// 랙·모듈은 새 표본이 왔을 때만 다시 계산 (PLC 주기마다 300개를 계산하지 않음)
IF NOT _bCalculated OR i_stState.nSampleSeq <> _nLastSeq OR q_bValid <> _bLastValid THEN
	_bCalculated := TRUE;
	_nLastSeq := i_stState.nSampleSeq;
	_bLastValid := q_bValid;
	_nOnlineRacks := 0;
	_bInitializing := FALSE;
	_bCharging := FALSE;
	_bDischarging := FALSE;
	_nBatWarn1 := 0;
	_nBatWarn2 := 0;
	FOR _nIndex := 1 TO 5 DO _anBatFault[_nIndex] := 0; END_FOR
	FOR _nRack := 1 TO GVL_PARAM.RACKS_PER_BMS DO
		q_astRack[_nRack] := _stRackEmpty;
		q_astRack[_nRack].DeviceIndex := (i_nDeviceIndex - 1) * UINT_TO_UDINT(GVL_PARAM.RACKS_PER_BMS) + UINT_TO_UDINT(_nRack);	// 전체 랙 순번 1부터
		q_astRack[_nRack].BatIndex := i_nDeviceIndex;
		q_astRack[_nRack].ModuleCount := UINT_TO_UDINT(i_stState.nModuleCount);
		q_astRack[_nRack].Status := 1; // b0 통신에러
		FOR _nModule := 1 TO GVL_PARAM.MODULES_PER_RACK DO
			_nIndex := (_nRack - 1) * GVL_PARAM.MODULES_PER_RACK + _nModule;
			q_astModule[_nIndex] := _stModuleEmpty;
			q_astModule[_nIndex].BatIndex := i_nDeviceIndex;
			q_astModule[_nIndex].RackIndex := UINT_TO_UDINT(_nRack);
			q_astModule[_nIndex].DeviceIndex := UINT_TO_UDINT(_nModule);
		END_FOR
		IF q_bValid AND _nRack <= i_stState.nRackCount THEN
			_nAnalog := (_nRack - 1) * 4;
			_nStatus := (_nRack - 1) * 9;
			_wOperation := i_stRaw.awRackStatus[_nStatus + 1];
			// 명세 RD-BAT-01 (v2.37): 배터리 eventMap v2. 칸 하나에 BMS 워드 2개 (첫 워드 b0~, 둘째 워드 b16~), 워드 안에서는 정의된 비트만 이어 붙임
			_wSysAlarm := i_stRaw.awRackStatus[_nStatus] AND SYS_ALARM_MASK;
			_wSysWarn := i_stRaw.awRackStatus[_nStatus + 2] AND SYS_WARN_MASK;
			_wSysError := i_stRaw.awRackStatus[_nStatus + 3] AND SYS_ERROR_MASK;
			_wModError := i_stRaw.awRackStatus[_nStatus + 4] AND MODULE_ERROR_MASK;
			_wErr1 := i_stRaw.awRackStatus[_nStatus + 5];
			_wErr2 := i_stRaw.awRackStatus[_nStatus + 6] AND ERROR_CODE2_MASK;
			_wFire := i_stRaw.awRackStatus[_nStatus + 7] AND FIRE_MASK;
			_wModule := i_stRaw.awRackStatus[_nStatus + 8] AND MODULE_STATUS_MASK;
			_wLock1 := 0;
			_wLock2 := 0;
			_wSelf1 := 0;
			_wSelf2 := 0;
			IF i_stState.abDetailValid[_nRack] THEN // 랙 상세는 순서대로 나눠 읽으므로 받은 랙만
				_wLock1 := i_stRaw.aawDetail[_nRack, 11] AND LOCK1_MASK;
				_wLock2 := i_stRaw.aawDetail[_nRack, 12] AND LOCK2_MASK;
				_wSelf1 := i_stRaw.aawDetail[_nRack, 13] AND SELF1_MASK;
				_wSelf2 := i_stRaw.aawDetail[_nRack, 14] AND SELF2_MASK;
			END_IF
			q_astRack[_nRack].Warning1 := WORD_TO_UDINT(_wSysWarn) OR SHL(WORD_TO_UDINT(_wSysAlarm), 16);	// S+2 | S+0
			// 명세 RD-BAT-01 (v2.48): 경고 비트 5개는 Warning2 b0~4 (S+4 b9 → b0, S+8 b0·2·4·6 → b1~4). '워드 2개' 규칙의 예외
			q_astRack[_nRack].Warning2 := WORD_TO_UDINT(SHR(_wModError, 9) AND 16#0001)
				OR SHL(WORD_TO_UDINT(_wModule AND 16#0001), 1)
				OR SHL(WORD_TO_UDINT(SHR(_wModule, 2) AND 16#0001), 2)
				OR SHL(WORD_TO_UDINT(SHR(_wModule, 4) AND 16#0001), 3)
				OR SHL(WORD_TO_UDINT(SHR(_wModule, 6) AND 16#0001), 4);
			// S+3 | S+4 (v2.48: b0~8 → b16~24, b10 → b25. b9는 Warning2)
			q_astRack[_nRack].Fault1 := WORD_TO_UDINT(_wSysError)
				OR SHL(WORD_TO_UDINT(_wModError AND 16#01FF), 16)
				OR SHL(WORD_TO_UDINT(SHR(_wModError, 10) AND 16#0001), 25);
			// S+7 (b0 → b0, b15 → b1) | S+8 (v2.48: b1·3·5·7·8 → b16~20. 경고 b0·2·4·6은 Warning2)
			q_astRack[_nRack].Fault2 := WORD_TO_UDINT(_wFire AND 16#0001) OR SHL(WORD_TO_UDINT(SHR(_wFire, 15)), 1)
				OR SHL(WORD_TO_UDINT(SHR(_wModule, 1) AND 16#0001), 16)
				OR SHL(WORD_TO_UDINT(SHR(_wModule, 3) AND 16#0001), 17)
				OR SHL(WORD_TO_UDINT(SHR(_wModule, 5) AND 16#0001), 18)
				OR SHL(WORD_TO_UDINT(SHR(_wModule, 7) AND 16#0001), 19)
				OR SHL(WORD_TO_UDINT(SHR(_wModule, 8) AND 16#0001), 20);
			// D+11 (b0·1 → b0·1, b3 → b2, b6~11 → b3~8) | D+12 (b0·1 → b16·17, b4~15 → b18~29)
			q_astRack[_nRack].Fault3 := WORD_TO_UDINT(_wLock1 AND 16#0003)
				OR SHL(WORD_TO_UDINT(SHR(_wLock1, 3) AND 16#0001), 2)
				OR SHL(WORD_TO_UDINT(SHR(_wLock1, 6) AND 16#003F), 3)
				OR SHL(WORD_TO_UDINT(_wLock2 AND 16#0003), 16)
				OR SHL(WORD_TO_UDINT(SHR(_wLock2, 4) AND 16#0FFF), 18);
			q_astRack[_nRack].Fault4 := WORD_TO_UDINT(_wErr1) OR SHL(WORD_TO_UDINT(_wErr2), 16);			// S+5 | S+6
			// D+13 | D+14 (b0~10 → b16~26, b12~15 → b27~30)
			q_astRack[_nRack].Fault5 := WORD_TO_UDINT(_wSelf1)
				OR SHL(WORD_TO_UDINT(_wSelf2 AND 16#07FF), 16)
				OR SHL(WORD_TO_UDINT(SHR(_wSelf2, 12) AND 16#000F), 27);
			_bRackWarn := (q_astRack[_nRack].Warning1 OR q_astRack[_nRack].Warning2) <> 0;	// v2.48: Warning2 포함
			_bRackFault := (q_astRack[_nRack].Fault1 OR q_astRack[_nRack].Fault2 OR q_astRack[_nRack].Fault3
				OR q_astRack[_nRack].Fault4 OR q_astRack[_nRack].Fault5) <> 0;
			_nBatWarn1 := _nBatWarn1 OR q_astRack[_nRack].Warning1;
			_nBatWarn2 := _nBatWarn2 OR q_astRack[_nRack].Warning2;
			_anBatFault[1] := _anBatFault[1] OR q_astRack[_nRack].Fault1;
			_anBatFault[2] := _anBatFault[2] OR q_astRack[_nRack].Fault2;
			_anBatFault[3] := _anBatFault[3] OR q_astRack[_nRack].Fault3;
			_anBatFault[4] := _anBatFault[4] OR q_astRack[_nRack].Fault4;
			_anBatFault[5] := _anBatFault[5] OR q_astRack[_nRack].Fault5;
			q_astRack[_nRack].Status := 0;
			q_astRack[_nRack].Status.1 := NOT _wOperation.0; // Initializing
			q_astRack[_nRack].Status.2 := _wOperation.3; // Ready = Idle RELAY ON
			q_astRack[_nRack].Status.3 := _wOperation.1; // Charge
			q_astRack[_nRack].Status.4 := _wOperation.2; // Discharge
			q_astRack[_nRack].Status.5 := _bRackWarn; // Warning 칸 중 하나라도 0이 아님
			q_astRack[_nRack].Status.6 := _bRackFault; // Fault 칸 중 하나라도 0이 아님
			q_astRack[_nRack].Status.7 := _wOperation.1 OR _wOperation.2 OR _wOperation.3; // Online
			q_astRack[_nRack].Status.10 := (SHR(i_stState.wRackContactor, _nRack - 1) AND 1) <> 0; // 랙 컨택터 붙음 (맵 v1.4 Input 27) [2026-11-13]
			q_astRack[_nRack].DcVoltage := WORD_TO_REAL(i_stRaw.awRackAnalog[_nAnalog]) * 0.1;
			q_astRack[_nRack].DcCurrent := F_UpsSignedWord(i_stRaw.awRackAnalog[_nAnalog + 1]) * 0.1;
			q_astRack[_nRack].Soc := WORD_TO_REAL(i_stRaw.awRackAnalog[_nAnalog + 2]) * 0.1;
			q_astRack[_nRack].Soh := WORD_TO_REAL(i_stRaw.awRackAnalog[_nAnalog + 3]);
			IF q_astRack[_nRack].Status.7 THEN _nOnlineRacks := _nOnlineRacks + 1; END_IF
			_bInitializing := _bInitializing OR NOT _wOperation.0;
			_bCharging := _bCharging OR _wOperation.1;
			_bDischarging := _bDischarging OR _wOperation.2;

			// 상세 데이터: 406칸. 모듈 슬롯 0부터 설치 수만큼 사용
			IF i_stState.abDetailValid[_nRack] THEN
				q_astRack[_nRack].MaxModuleTemp := F_UpsSignedWord(i_stRaw.aawDetail[_nRack, 0]) * 0.1;
				q_astRack[_nRack].MinModuleTemp := F_UpsSignedWord(i_stRaw.aawDetail[_nRack, 1]) * 0.1;
				q_astRack[_nRack].AvgModuleTemp := F_UpsSignedWord(i_stRaw.aawDetail[_nRack, 2]) * 0.1;
				q_astRack[_nRack].MaxCellVoltage := WORD_TO_REAL(i_stRaw.aawDetail[_nRack, 3]) * 0.001;
				q_astRack[_nRack].MinCellVoltage := WORD_TO_REAL(i_stRaw.aawDetail[_nRack, 4]) * 0.001;
				q_astRack[_nRack].AvgCellVoltage := WORD_TO_REAL(i_stRaw.aawDetail[_nRack, 5]) * 0.001;
				_wCellMax := 0;
				_wCellMin := 16#FFFF;
				_fTempMax := -1.0E6;
				_fTempMin := 1.0E6;
				FOR _nModule := 1 TO MIN(i_stState.nModuleCount, GVL_PARAM.MODULES_PER_RACK) DO
					_nIndex := (_nRack - 1) * GVL_PARAM.MODULES_PER_RACK + _nModule;
					// @MAP 랙 상세 D+15+m (첫 랙 30516부터), uint16 x0.01 V. m = 모듈 번호 - 1
					q_astModule[_nIndex].ModuleVolatge1 := WORD_TO_REAL(i_stRaw.aawDetail[_nRack, 14 + _nModule]) * 0.01;
					// ModuleVolatge2/3은 BMS 맵에 없어 _stModuleEmpty의 0 유지
					_fTemp := F_UpsSignedWord(i_stRaw.aawDetail[_nRack, 31 + _nModule]) * 0.1; // 맵은 모듈당 최고 온도 1개
					q_astModule[_nIndex].ModuleTemp1 := _fTemp;
					IF _fTemp > _fTempMax THEN
						_fTempMax := _fTemp;
						q_astRack[_nRack].MaxModuleTempLocationFromModule := UINT_TO_UDINT(_nModule);
					END_IF
					IF _fTemp < _fTempMin THEN
						_fTempMin := _fTemp;
						q_astRack[_nRack].MinModuleTempLocationFromModule := UINT_TO_UDINT(_nModule);
					END_IF
					_pCell := ADR(q_astModule[_nIndex].CellVoltage1);
					FOR _nCell := 1 TO MIN(GVL_PARAM.CELLS_PER_MODULE, 20) DO	// 설치 셀 수만 (맵은 모듈당 20칸, 레코드 CellVoltage15~20은 0으로 남음)
						_wCell := i_stRaw.aawDetail[_nRack, 66 + 20 * (_nModule - 1) + _nCell - 1];
						_pCell[_nCell - 1] := WORD_TO_REAL(_wCell) * 0.001;
						IF _wCell > _wCellMax THEN
							_wCellMax := _wCell;
							q_astRack[_nRack].MaxCellVoltageLocationFromModule := UINT_TO_UDINT(_nModule);
							q_astRack[_nRack].MaxCellVoltageLocationFromCell := UINT_TO_UDINT(_nCell);
						END_IF
						IF _wCell < _wCellMin THEN
							_wCellMin := _wCell;
							q_astRack[_nRack].MinCellVoltageLocationFromModule := UINT_TO_UDINT(_nModule);
							q_astRack[_nRack].MinCellVoltageLocationFromCell := UINT_TO_UDINT(_nCell);
						END_IF
					END_FOR
				END_FOR
			END_IF
		END_IF
	END_FOR
END_IF

IF q_bValid THEN
	q_stBat.OnlineRackCount := _nOnlineRacks;
	q_stBat.Status := 0;
	q_stBat.Status.1 := _bInitializing;
	q_stBat.Status.2 := NOT _bInitializing AND _nOnlineRacks = 0; // Standby
	q_stBat.Status.3 := _nOnlineRacks > 0 AND NOT _bCharging AND NOT _bDischarging; // Ready
	q_stBat.Status.4 := _bCharging;
	q_stBat.Status.5 := _bDischarging;
	// 명세 RD-BAT-02 (v2.48): BAT Warning1·Warning2·Fault1~5 = 랙 값 OR (칸 배치는 RACK과 같음). 나머지 칸은 0
	q_stBat.Warning1 := _nBatWarn1;
	q_stBat.Warning2 := _nBatWarn2;
	q_stBat.Fault1 := _anBatFault[1];
	q_stBat.Fault2 := _anBatFault[2];
	q_stBat.Fault3 := _anBatFault[3];
	q_stBat.Fault4 := _anBatFault[4];
	q_stBat.Fault5 := _anBatFault[5];
	q_stBat.Status.6 := (_nBatWarn1 OR _nBatWarn2) <> 0;	// v2.48: Warning2 포함
	q_stBat.Status.7 := (_anBatFault[1] OR _anBatFault[2] OR _anBatFault[3] OR _anBatFault[4] OR _anBatFault[5]) <> 0;
	q_stBat.Status.9 := i_stState.bSystemLock; // Emergency = 어느 랙이든 System Lock (Level 3, 현장 해제 필요)
	q_stBat.Status.11 := i_stState.bChargeContactorClosed; // 충전 컨택터 붙음 (맵 v1.4 Input 26 b0) [2026-11-13]
	q_stBat.Status.12 := i_stState.bDischargeContactorClosed; // 방전 컨택터 붙음 (맵 v1.4 Input 26 b1) [2026-11-13]
	q_stBat.Status.13 := i_stState.wRackContactor <> 0; // 명세 RD-BAT-02 (v2.28): 랙 컨택터 닫힘 = 랙 하나라도 닫힘 (Input 27 ≠ 0, EMS 단선도 DC 컨택터)
	// b8 Balancing, b10 E-stop은 맵에 정보가 없어 항상 0 (미지원)
END_IF
// Eol, 랙 충·방전 제한, 온도 셀 위치는 맵에 없어 0. RACK b8 Precharge·b9 Balancing은 미지원이라 0.

END_FUNCTION_BLOCK

// ---- 20_Module/Ups/F_UpsSignedWord.TcPOU
FUNCTION F_UpsSignedWord : REAL
VAR_INPUT i_wRaw : WORD; END_VAR

IF i_wRaw >= 16#8000 THEN
	F_UpsSignedWord := DINT_TO_REAL(WORD_TO_DINT(i_wRaw) - 65536);
ELSE
	F_UpsSignedWord := WORD_TO_REAL(i_wRaw);
END_IF

END_FUNCTION

// ---- 20_Module/Report/FB_RptSebangUps.TcPOU
FUNCTION_BLOCK FB_RptSebangUps // UPS 계측값 → UPS 보고값
VAR_INPUT
	i_stState : ST_UpsState; // 장비 상태
	i_nDeviceIndex : UDINT; // UPS 번호
	i_nOperationMode : UDINT := 1; // 0 수동, 1 자동 (FB_UpsCommand.q_nOperationMode)
END_VAR
VAR_OUTPUT
	q_stUps : ST_UpsPublish_V1; // UPS 보고값
	q_bValid : BOOL; // 유효한 장비 데이터
END_VAR
VAR
	_stEmpty : ST_UpsPublish_V1;
	_awWarn : ARRAY[0..7] OF WORD; // 워드별 경고장 비트 (I44~I51)
	_awFault : ARRAY[0..7] OF WORD; // 워드별 중고장 비트 (I44~I51)
	_i : INT;
	_b : INT; // 워드 안 비트 번호
	_wBit : WORD;
	_nWarnPos : INT; // 다음에 채울 Warning1 비트
	_nFault1Pos : INT; // 다음에 채울 Fault1 비트
	_nFault2Pos : INT; // 다음에 채울 Fault2 비트
END_VAR
VAR CONSTANT
	// 세방 맵 v3.2 Alarm Flag 색. 순서 = I44 입력, I45 정류부, I46 BBC, I47 출력, I48 인버터, I49 바이패스, I50 STATUS1, I51 STATUS2
	WARN_MASK : ARRAY[0..7] OF WORD := [16#0700, 16#0003, 16#0007, 16#00FF, 16#0000, 16#03FF, 16#0000, 16#0701]; // 경고장(노랑)
	FAULT_MASK : ARRAY[0..7] OF WORD := [16#F8FF, 16#667C, 16#0FB8, 16#3F00, 16#803F, 16#0000, 16#0081, 16#7800]; // 중고장(주황)
	FAULT1_LAST_WORD : INT := 2; // 중고장 I44~I46 → Fault1, I47~I51 → Fault2 (회사 eventMap)
END_VAR

q_stUps := _stEmpty;
q_stUps.DeviceIndex := i_nDeviceIndex;
q_stUps.Status := 1; // b0 통신에러
q_bValid := i_stState.bValid;
IF NOT q_bValid THEN
	RETURN;
END_IF

// 명세 RD-UPS-02 (v2.20, 회사 eventMap '001.UPS 경고장비트맵'): 마스크로 거른 경고장·중고장 비트를
// 맵 워드 순서(I44→I51), 워드 안 비트 순서로 b0부터 빈칸 없이 채운다. 마스크 밖 비트(운전 상태·예약)는 버림
//   Warning1 = 경고장 30개 (I44·I45·I46·I47·I49·I51) b0~b29, Warning2·3 = 0
//   Fault1 = I44·I45·I46 중고장 30개 b0~b29, Fault2 = I47·I48·I50·I51 중고장 19개 b0~b18, Fault3 = 0
// 마스크가 바뀌면 그 뒤 비트 자리가 모두 밀리므로 eventMap도 같이 고쳐야 함
_nWarnPos := 0;
_nFault1Pos := 0;
_nFault2Pos := 0;
FOR _i := 0 TO 7 DO
	_awWarn[_i] := i_stState.awAlarmStatus[_i] AND WARN_MASK[_i];
	_awFault[_i] := i_stState.awAlarmStatus[_i] AND FAULT_MASK[_i];
	FOR _b := 0 TO 15 DO
		_wBit := SHL(WORD#1, _b);
		IF (WARN_MASK[_i] AND _wBit) <> 0 THEN
			IF (_awWarn[_i] AND _wBit) <> 0 THEN
				q_stUps.Warning1 := q_stUps.Warning1 OR SHL(UDINT#1, _nWarnPos);
			END_IF
			_nWarnPos := _nWarnPos + 1;
		END_IF
		IF (FAULT_MASK[_i] AND _wBit) <> 0 THEN
			IF _i <= FAULT1_LAST_WORD THEN
				IF (_awFault[_i] AND _wBit) <> 0 THEN
					q_stUps.Fault1 := q_stUps.Fault1 OR SHL(UDINT#1, _nFault1Pos);
				END_IF
				_nFault1Pos := _nFault1Pos + 1;
			ELSE
				IF (_awFault[_i] AND _wBit) <> 0 THEN
					q_stUps.Fault2 := q_stUps.Fault2 OR SHL(UDINT#1, _nFault2Pos);
				END_IF
				_nFault2Pos := _nFault2Pos + 1;
			END_IF
		END_IF
	END_FOR
END_FOR

// 명세 RD-UPS-01: 상태 칸 (인터페이스 08.UPS 2026-11-12). 맵 워드: I45 정류부, I46 BBC, I48 인버터, I50 STATUS1, I51 STATUS2
// 운전 모드 (2026-11-25): EMS UPS 명령 101 수동·102 자동을 반영. SystemOperationMode는 0 유지
q_stUps.SystemOperationMode := 0;
q_stUps.OperationMode := i_nOperationMode;
q_stUps.Status := 0;
q_stUps.Status.1 := (q_stUps.Warning1 OR q_stUps.Warning2 OR q_stUps.Warning3) <> 0; // 경고 있음
q_stUps.Status.2 := (q_stUps.Fault1 OR q_stUps.Fault2 OR q_stUps.Fault3) <> 0; // 고장 있음
q_stUps.Status.3 := i_stState.bEmergencyStop; // e-stop (I50 b0)
q_stUps.Status.4 := i_stState.wStatus1.13; // 충전 중 (I50 b13 Batt charg Flag)

q_stUps.UPS_ModeStatus := 0;
q_stUps.UPS_ModeStatus.0 := i_stState.nBatMode = 0; // 부동충전 (BAT Mode 값을 비트로 나눔)
q_stUps.UPS_ModeStatus.1 := i_stState.nBatMode = 1; // 균등충전
q_stUps.UPS_ModeStatus.2 := i_stState.nBatMode = 2; // 대기
q_stUps.UPS_ModeStatus.3 := i_stState.nBatMode = 3; // 주기적 방전
q_stUps.UPS_ModeStatus.4 := i_stState.nBatMode = 4; // 펄스 방전
q_stUps.UPS_ModeStatus.5 := i_stState.nBatMode = 5; // 간헐충전
q_stUps.UPS_ModeStatus.6 := i_stState.wRectAlarm.8; // 비상 방전 (I45 b8 Regen mode)
q_stUps.UPS_ModeStatus.7 := i_stState.bTemperatureEnabled; // 온도보상충전 (I51 b2, 다른 모드와 동시 가능)
q_stUps.UPS_ModeStatus.8 := i_stState.wInverterAlarm.7; // ECO 모드 (I48 b7)
q_stUps.UPS_ModeStatus.9 := i_stState.wStatus1.12; // PRLT 모드 (I50 b12)
q_stUps.UPS_ModeStatus.10 := i_stState.wStatus1.11; // Droop 모드 (I50 b11)
q_stUps.UPS_ModeStatus.11 := i_stState.wRectAlarm.15; // VSM 모드 (I45 b15)
q_stUps.UPS_ModeStatus.12 := i_stState.wRectAlarm.8; // Regen 모드 (I45 b8, b6과 같은 비트)

q_stUps.MCCB_Status := SHR(WORD_TO_UDINT(i_stState.wStatus1), 1) AND 16#3F; // I50 b1~b6 → b0~b5 (b5 Out C/B는 1이 개방)
q_stUps.MCCB_Status.6 := i_stState.wOpCode.3; // 배터리 MCCB Trip (H11 OP-CODE b3, 1 = Trip, 세방 회신 2026-11-25, 명세 RD-UPS-01 v2.50)

q_stUps.RectStatus := 0;
q_stUps.RectStatus.0 := i_stState.bRectOn; // 정류부 기동 (I45 b11)
q_stUps.RectStatus.1 := i_stState.bRectNormal; // 정류부 정상 (I45 b12)
q_stUps.RectStatus.2 := i_stState.wRectAlarm.8; // Regen (I45 b8, 비상 방전)

q_stUps.BBCStatus := 0;
q_stUps.BBCStatus.0 := i_stState.bBbcOn; // 배터리 컨버터 기동 (I46 b12)
q_stUps.BBCStatus.1 := i_stState.bBbcNormal; // 배터리 컨버터 정상 (I46 b13)

q_stUps.InverterStatus := 0;
q_stUps.InverterStatus.0 := i_stState.bInverterOn; // 인버터 기동 (I48 b6)
q_stUps.InverterStatus.1 := i_stState.bInverterNormal; // 인버터 정상 (I48 b14)
q_stUps.InverterStatus.2 := i_stState.bOnInverter; // 인버터 출력 (I48 b13)

q_stUps.BypassStatus := 0;
q_stUps.BypassStatus.0 := i_stState.bOnBypass; // 바이패스 출력 (I48 b12)

q_stUps.LineInputVoltage_R := i_stState.fInputVoltageRV;
q_stUps.LineInputVoltage_S := i_stState.fInputVoltageSV;
q_stUps.LineInputVoltage_T := i_stState.fInputVoltageTV;
q_stUps.InputFrequency := i_stState.fInputFrequencyHz;
q_stUps.InputCurrent_R := i_stState.fInputCurrentRA;
q_stUps.InputCurrent_S := i_stState.fInputCurrentSA;
q_stUps.InputCurrent_T := i_stState.fInputCurrentTA;
q_stUps.InverterVoltage_R := i_stState.fInverterVoltageRV;
q_stUps.InverterVoltage_S := i_stState.fInverterVoltageSV;
q_stUps.InverterVoltage_T := i_stState.fInverterVoltageTV;
q_stUps.InverterCurrent_R := i_stState.fInverterCurrentRA;
q_stUps.InverterCurrent_S := i_stState.fInverterCurrentSA;
q_stUps.InverterCurrent_T := i_stState.fInverterCurrentTA;
q_stUps.BypassLineVoltage_R := i_stState.fBypassVoltageRV;
q_stUps.BypassLineVoltage_S := i_stState.fBypassVoltageSV;
q_stUps.BypassLineVoltage_T := i_stState.fBypassVoltageTV;
q_stUps.BypassFrequency := i_stState.fBypassFrequencyHz;
q_stUps.LineOutputVoltage_R := i_stState.fOutputVoltageRV;
q_stUps.LineOutputVoltage_S := i_stState.fOutputVoltageSV;
q_stUps.LineOutputVoltage_T := i_stState.fOutputVoltageTV;
q_stUps.FrequencyOutput := i_stState.fOutputFrequencyHz;
q_stUps.OutputCurrent_R := i_stState.fOutputCurrentRA;
q_stUps.OutputCurrent_S := i_stState.fOutputCurrentSA;
q_stUps.OutputCurrent_T := i_stState.fOutputCurrentTA;
q_stUps.DcLinkVoltage := i_stState.fDcLinkVoltageV;
q_stUps.DcLinkVoltage_High := i_stState.fDcLinkHighVoltageV;
q_stUps.DcLinkVoltage_Low := i_stState.fDcLinkLowVoltageV;
q_stUps.BatteryVoltage := i_stState.fBatteryVoltageV;
q_stUps.BatteryCurrent := i_stState.fBatteryCurrentA;
q_stUps.MPI_A_Current := i_stState.fMpiCurrentAA;
q_stUps.MPI_B_Current := i_stState.fMpiCurrentBA;
q_stUps.MPI_C_Current := i_stState.fMpiCurrentCA;
q_stUps.InputApparentPower := i_stState.fInputApparentPowerKva;
q_stUps.OutputApparentPower := i_stState.fOutputApparentPowerKva;
q_stUps.OutputActivePower := i_stState.fOutputActivePowerKw;
q_stUps.Temp1 := i_stState.fTemperature1C;
q_stUps.Temp2 := i_stState.fTemperature2C;
q_stUps.Temp3 := i_stState.fTemperature3C;
q_stUps.Temp4 := i_stState.fTemperature4C;
q_stUps.Temp5 := i_stState.fTemperature5C;
q_stUps.Temp6 := i_stState.fBatteryRoomTemperatureC;

END_FUNCTION_BLOCK

// ---- 20_Module/Report/FB_RptLsImd1000.TcPOU
FUNCTION_BLOCK FB_RptLsImd1000		// LS IMD1000 읽은 값 → IMD 보고값 (인터페이스\22. IMD.xlsx)
(* 2026-11-09. 명세 DV-11·RD-IMD-01 (v1.8)
   Status (사용자 결정 2026-11-09, 저항이 높은 경보부터)
     b0 통신에러 = 통신 이상 또는 아직 못 읽음 (나머지 칸 0)
     b1 Pre-Warning = Pre Alarm#3 동작 (IR 210 b3, 초기값 100 kΩ)
     b2 Warning = Pre Alarm#1 OR #2 동작 (IR 210 b1·b2, 초기값 40·70 kΩ)
     b3 Fault = 자가진단 오류 (IR 209 b0~2 메모리·RTC·교정) OR Device 이상 (IR 211 b1)
     b4 Alarm = Ins. Alarm 동작 (IR 210 b0, 초기값 10 kΩ)
     b5 Internal test = Self Test 진행 중 (IR 215 = 1)
     b6 External test = 버튼·DI Self Test 입력 (IR 206 b0·b1)
   Fault1 b0 = System 연결 이상 (IR 211 b2), b1 = PE 연결 이상 (IR 211 b0)
   PreAlarmSettingValue = Pre Alarm#1 Pick-up, MainAlarmSettingValue = Ins. Alarm Pick-up (설정 영역을 못 읽었으면 0)
   DeviceErrorLocation·InsulationResistanceFaultLocation은 Bender 항목이라 0 *)
VAR_INPUT
	i_stState		: ST_LsImd1000State;	// 장비 상태 (FB_LsImd1000.q_stState)
	i_nDeviceIndex	: UDINT;				// IMD 번호 (1부터)
END_VAR
VAR_OUTPUT
	q_stImd			: ST_ImdPublish_V1;		// IMD 보고값
	q_bValid		: BOOL;					// 유효한 장비 데이터
END_VAR
VAR
	_stEmpty		: ST_ImdPublish_V1;
END_VAR

q_stImd := _stEmpty;
q_stImd.DeviceIndex := i_nDeviceIndex;
q_stImd.Status := 1;	// b0 통신에러
q_bValid := i_stState.bValid;
IF NOT q_bValid THEN
	RETURN;
END_IF

q_stImd.Status := 0;
q_stImd.Status.1 := i_stState.wAlarm.3;
q_stImd.Status.2 := i_stState.wAlarm.1 OR i_stState.wAlarm.2;
q_stImd.Status.3 := (i_stState.wSelfDiag AND 16#0007) <> 0 OR i_stState.wConnect.1;
q_stImd.Status.4 := i_stState.wAlarm.0;
q_stImd.Status.5 := i_stState.wSelfTest = 1;
q_stImd.Status.6 := i_stState.wDiState.0 OR i_stState.wDiState.1;

q_stImd.InsulationResistance := i_stState.fInsulation;
IF i_stState.bSetValid THEN
	q_stImd.PreAlarmSettingValue := i_stState.nPre1Pickup;
	q_stImd.MainAlarmSettingValue := i_stState.nInsPickup;
END_IF
q_stImd.Fault1.0 := i_stState.wConnect.2;
q_stImd.Fault1.1 := i_stState.wConnect.0;

END_FUNCTION_BLOCK

// ---- 20_Module/Report/FB_RptTempHum.TcPOU
FUNCTION_BLOCK FB_RptTempHum		// 온습도계 읽은 값 → 온도 보고값 (인터페이스\07.Temperature Sensor.xlsx, 토픽 temperature_sensor)
(* 2026-11-09. status b0 통신에러(통신 이상·값 무효면 1, 온도·습도 0). location은 설치 위치 번호
   (1 PCS실, 2 BAT실, 3 UPS실, 4 FC 컨테이너실, 5 외부) *)
VAR_INPUT
	i_stState		: ST_TempHumState;		// 장비 상태 (드라이버 q_stState)
	i_nDeviceIndex	: UDINT;				// 장치 번호 (0부터, 기존 temperature_sensor 시험 데이터와 같음)
	i_nLocation		: UDINT;				// 설치 위치
END_VAR
VAR_OUTPUT
	q_stTemp		: ST_TempPublish_V1;	// 보고값
	q_bValid		: BOOL;					// 유효한 장비 데이터
END_VAR
VAR
	_stEmpty		: ST_TempPublish_V1;
END_VAR

q_stTemp := _stEmpty;
q_stTemp.DeviceIndex := i_nDeviceIndex;
q_stTemp.location := i_nLocation;
q_stTemp.status := 1;	// b0 통신에러
q_bValid := i_stState.bValid;
IF NOT q_bValid THEN
	RETURN;
END_IF
q_stTemp.status := 0;
q_stTemp.temperature := i_stState.fTemp;
q_stTemp.humidity := i_stState.fHum;

END_FUNCTION_BLOCK

// ---- 20_Module/Driver/Esolution/FB_BmsRackCommand.TcPOU
FUNCTION_BLOCK FB_BmsRackCommand		// BMS 랙 컨택터 개별 제어: EMS 랙 명령 → 랙 선택표(BMS 40001 랙 비트) 갱신 요청
(* 2026-11-10. 명세 WR-BAT-01 (v2.5). 인터페이스 100.Command BAT CommandType 11 랙 닫기 / 12 랙 열기 (Value = 랙 번호)
   BAT 질의 Q4 답변: 랙 개별·일괄 제어 모두 지원. 일괄은 CommandType 1·2 (시스템 컨택터 40013, 기존 코어 경로)
   - 랙 선택표(비트 n-1 = 랙 n, 1 = 사용)를 기억하고, 명령마다 그 랙 비트만 바꾼 표 전체를 BMS에 쓰게 한다
   - 장비 쓰기는 하지 않는다. q_bWriteReq·q_wWriteMask를 MAIN이 보고 드라이버 M_SetRackMask를 부르고 결과를 돌려준다
   - 선택표는 PERSISTENT (i_wRestore로 시작 때 한 번 읽고, q_wMask를 MAIN이 저장). 저장값이 없으면(0) 설치된 랙 전부
   - 거절: 랙 번호 범위 밖(BadRequest), 마지막 남은 랙 열기(BadRequest: 0이면 BMS가 전 랙 사용 안 함 → 전체는 일괄 2 열기로)
   - 드라이버가 바쁘면(Busy) WRITE_TIMEOUT 동안 다시 시도. 그 밖의 거절(쓰기 막힘, 통신 불가 등)은 바로 그 결과로 끝
   - 같은 상태로 바꾸는 명령도 표 전체를 다시 씀 (BMS가 다시 켜져 표가 달라졌을 때 맞춤)
   - [2026-11-13] BMS 맵 v1.4 랙 컨택터 상태(Input 30027)를 받으면 그 실제 상태를 바탕으로 비트를 바꿈.
     40013(랙 전체 연결)으로 다 붙은 뒤 옛 선택표로 써서 다른 랙을 떼는 일을 막음. 상태가 없으면 기억한 선택표 *)
VAR_INPUT
	i_stCmd			: ST_BatRackCmd;	// EMS 랙 명령 (번호가 바뀌면 새 명령)
	i_nRackCount	: UINT;				// 설치된 랙 수 (GVL_PARAM.RACKS_PER_BMS)
	i_wRestore		: WORD;				// 처음 호출 때 한 번 읽는 저장된 선택표 (GVL_PERSIST.g_awBmsRackMask[n])
	i_bAccepted		: BOOL;				// 지난 스캔의 쓰기 요청을 드라이버가 받음 (M_SetRackMask 반환값)
	i_eDriverResult	: E_UpsResult;		// 지난 스캔 드라이버 결과 (q_eRequestResult). 요청하지 않은 스캔은 None
	i_wActual		: WORD;				// BMS 랙 컨택터 실제 상태 (q_stState.wRackContactor, 30027) [2026-11-13]
	i_bActualValid	: BOOL;				// i_wActual을 믿을 수 있음 (q_stState.bContactorFeedbackKnown)
END_VAR
VAR_OUTPUT
	q_wMask			: WORD;				// 지금 선택표 (드라이버가 받은 값). MAIN이 GVL_PERSIST에 씀
	q_bMaskChanged	: BOOL;				// 이 스캔에 q_wMask가 바뀜 (PERSISTENT 바로 저장 요청)
	q_bWriteReq		: BOOL;				// 드라이버에 쓰기 요청 중
	q_wWriteMask	: WORD;				// 쓸 선택표
	q_eResult		: E_UpsResult;		// 마지막 명령 결과
	q_nLastSeq		: UDINT;			// 마지막으로 처리한 명령 번호
END_VAR
VAR
	_bInit			: BOOL;
	_wInstalled		: WORD;
	_wNew			: WORD;
	_wOld			: WORD;
	_wBase			: WORD;				// 바꿀 바탕 (실제 상태 또는 기억한 선택표)
	_tonWait		: TON;
END_VAR
VAR CONSTANT
	WRITE_TIMEOUT	: TIME := T#5S;		// 드라이버가 바쁠 때 다시 시도하는 시간
END_VAR

q_bMaskChanged := FALSE;
_wInstalled := SHL(WORD#1, MIN(i_nRackCount, 16)) - 1;
IF NOT _bInit THEN
	q_wMask := i_wRestore AND _wInstalled;
	IF q_wMask = 0 THEN
		q_wMask := _wInstalled;	// 저장값 없음 → 설치된 랙 전부
	END_IF
	_bInit := TRUE;
END_IF
_wOld := q_wMask;

// 1) 지난 스캔 쓰기 요청의 결과
IF q_bWriteReq THEN
	_tonWait(IN := TRUE, PT := WRITE_TIMEOUT);
	IF i_bAccepted THEN
		q_wMask := q_wWriteMask;
		q_eResult := E_UpsResult.Accepted;
		q_bWriteReq := FALSE;
	ELSIF i_eDriverResult <> E_UpsResult.None AND i_eDriverResult <> E_UpsResult.Busy THEN
		q_eResult := i_eDriverResult;	// 쓰기 막힘, 통신 불가, 설정 오류 등
		q_bWriteReq := FALSE;
	ELSIF _tonWait.Q THEN
		q_eResult := E_UpsResult.Busy;	// 계속 바빠서 포기
		q_bWriteReq := FALSE;
	END_IF
	IF NOT q_bWriteReq THEN
		_tonWait(IN := FALSE);
	END_IF
END_IF

// 2) 새 명령 (처리 중인 요청이 있으면 그것을 버리고 새 명령으로)
IF i_stCmd.nSeq <> q_nLastSeq AND i_stCmd.nSeq <> 0 THEN
	q_nLastSeq := i_stCmd.nSeq;
	q_bWriteReq := FALSE;
	_tonWait(IN := FALSE);
	IF i_stCmd.nRack < 1 OR i_stCmd.nRack > i_nRackCount OR i_stCmd.nRack > 16 THEN
		q_eResult := E_UpsResult.BadRequest;
	ELSE
		IF i_bActualValid THEN
			_wBase := i_wActual AND _wInstalled;	// 실제 상태 바탕
		ELSE
			_wBase := q_wMask;
		END_IF
		IF i_stCmd.bClose THEN
			_wNew := _wBase OR SHL(WORD#1, i_stCmd.nRack - 1);
		ELSE
			_wNew := _wBase AND NOT SHL(WORD#1, i_stCmd.nRack - 1);
		END_IF
		IF _wNew = 0 THEN
			q_eResult := E_UpsResult.BadRequest;	// 마지막 랙: 전체 열기는 일괄 명령(2)으로
		ELSE
			q_wWriteMask := _wNew;
			q_bWriteReq := TRUE;
			q_eResult := E_UpsResult.None;	// 처리 중
		END_IF
	END_IF
END_IF

q_bMaskChanged := q_wMask <> _wOld;

END_FUNCTION_BLOCK

// ---- 20_Module/Driver/Esolution/FB_BmsContactorCommand.TcPOU
FUNCTION_BLOCK FB_BmsContactorCommand		// BMS 컨택터 하나씩 제어: EMS 명령 번호 5~10 → 드라이버 M_SetControl 요청
(* 2026-11-13. 인터페이스 100.Command BAT CommandType 5~10, BMS 맵 v1.4 Holding 40013~40015
   5 시스템(랙 전체 40013) 연결   6 시스템 차단
   7 충전 컨택터(40014) 닫기      8 충전 컨택터 열기
   9 방전 컨택터(40015) 닫기      10 방전 컨택터 열기
   3 비상정지 (40012 Emergency Shutdown = 1). 2026-11-23 명세 v2.33: 코어(F_BatCmdAllowed)가 지령원 EStop을 거절해 이쪽으로 옮김
   4 초기화 (40031 Reset System = 1, 비상차단 해제). 2026-11-23 명세 v2.34 (O-19 A)
   - 장비 쓰기는 하지 않는다. q_bWriteReq·q_eControl·q_bOn을 MAIN이 보고 드라이버 M_SetControl을 부르고 결과를 돌려준다
   - 3~10 밖이면 BadRequest. 드라이버가 바쁘면(Busy) WRITE_TIMEOUT 동안 다시 시도. 그 밖의 거절(쓰기 막힘, 통신 불가 등)은 바로 그 결과로 끝
   - 코어 순서(유닛 정지 확인)는 거치지 않는다 (랙 개별 11·12와 같음). 일괄 투입·개방은 1·2 (코어 경로) *)
VAR_INPUT
	i_stCmd			: ST_BatCtlCmd;		// EMS 명령 (번호가 바뀌면 새 명령)
	i_bAccepted		: BOOL;				// 지난 스캔의 쓰기 요청을 드라이버가 받음 (M_SetControl 반환값)
	i_eDriverResult	: E_UpsResult;		// 지난 스캔 드라이버 결과 (q_eRequestResult). 요청하지 않은 스캔은 None
END_VAR
VAR_OUTPUT
	q_bWriteReq		: BOOL;				// 드라이버에 쓰기 요청 중
	q_eControl		: E_EsolutionControl;	// 쓸 컨택터
	q_bOn			: BOOL;				// TRUE = 닫기(붙이기), FALSE = 열기(떼기)
	q_eResult		: E_UpsResult;		// 마지막 명령 결과
	q_nLastSeq		: UDINT;			// 마지막으로 처리한 명령 번호
END_VAR
VAR
	_tonWait		: TON;
END_VAR
VAR CONSTANT
	WRITE_TIMEOUT	: TIME := T#5S;		// 드라이버가 바쁠 때 다시 시도하는 시간
END_VAR

// 1) 지난 스캔 쓰기 요청의 결과
IF q_bWriteReq THEN
	_tonWait(IN := TRUE, PT := WRITE_TIMEOUT);
	IF i_bAccepted THEN
		q_eResult := E_UpsResult.Accepted;
		q_bWriteReq := FALSE;
	ELSIF i_eDriverResult <> E_UpsResult.None AND i_eDriverResult <> E_UpsResult.Busy THEN
		q_eResult := i_eDriverResult;	// 쓰기 막힘, 통신 불가 등
		q_bWriteReq := FALSE;
	ELSIF _tonWait.Q THEN
		q_eResult := E_UpsResult.Busy;	// 계속 바빠서 포기
		q_bWriteReq := FALSE;
	END_IF
	IF NOT q_bWriteReq THEN
		_tonWait(IN := FALSE);
	END_IF
END_IF

// 2) 새 명령 (처리 중인 요청이 있으면 그것을 버리고 새 명령으로)
IF i_stCmd.nSeq <> q_nLastSeq AND i_stCmd.nSeq <> 0 THEN
	q_nLastSeq := i_stCmd.nSeq;
	q_bWriteReq := FALSE;
	_tonWait(IN := FALSE);
	q_eResult := E_UpsResult.None;	// 처리 중
	CASE i_stCmd.nType OF
		3:		q_eControl := E_EsolutionControl.EmergencyShutdown;
		4:		q_eControl := E_EsolutionControl.ResetSystem;
		5, 6:	q_eControl := E_EsolutionControl.SystemContactor;
		7, 8:	q_eControl := E_EsolutionControl.ChargeContactor;
		9, 10:	q_eControl := E_EsolutionControl.DischargeContactor;
	ELSE
		q_eResult := E_UpsResult.BadRequest;
	END_CASE
	IF q_eResult = E_UpsResult.None THEN
		q_bOn := (i_stCmd.nType MOD 2) = 1 OR i_stCmd.nType = 4;	// 3 비상정지·4 초기화 = 켜기(1), 5·7·9 = 닫기
		q_bWriteReq := TRUE;
	END_IF
END_IF

END_FUNCTION_BLOCK

// ---- 20_Module/Ups/FB_UpsSafetyResponse.TcPOU
FUNCTION_BLOCK FB_UpsSafetyResponse		// 사고·고장 대응 동작 (C안): 원인 → UPS·BMS 명령, 될 때까지 2초마다 다시 보내고 10초 넘으면 오류 표시
(* 2026-11-17. 명세 SQ-05 (v2.16), 동작시퀀스 7쪽 표. 기반 없음(신규).
   변경: 2026-11-18 ESD(b12) 대응을 나눔: 바이패스 절체 빼고 인버터 정지(H105) 추가, 순서 기다리지 않고 연달아 보냄 (명세 v2.18)
   변경: 2026-11-20 화재(b11)는 ESD처럼: 바이패스 절체 안 함, 인버터·BBC·정류부를 기다리지 않고 연달아 (명세 SQ-05 v2.31)
   변경: 2026-11-20 바이패스 이상(UPS Warning1 b16~25 = I49)이고 아직 바이패스가 아니면 바이패스 절체를 보내지 않음 → q_bBypassBlocked (v2.31, O-17)
   변경: 2026-11-20 세방 맵 '인버터정지 To Bypass': 출력·인버터 중고장, 화재, MBS C/B Fail(대응 원인 b13)은 바이패스 절체가
         확인된 뒤 인버터 정지(H105)도 보냄. 절체가 확인 안 되면 인버터를 끄지 않음(부하 유지). 원인은 q_nRespCause (명세 SQ-05 v2.30)
   변경: 2026-11-18 "3초 확인·최대 3번 → 실패로 멈춤"을 "될 때까지 2초마다 계속 보냄, 10초 넘게 안 되면 오류 표시(그 뒤에도 계속)"로 바꿈 (명세 v2.19, 데스틴 PCS 통신 방식)
   - 원인은 FB_UpsSafetyStage.q_nRespCause (지금 걸린 대응 원인, v2.30). 여러 원인이면 동작을 합친다
   - 동작 6개 (비트): 0 충전 컨택터 열기(BMS 40014=0), 1 BMS 컨택터 전부 열기(40013~15=0),
     2 바이패스 절체(UPS H109), 3 BBC 정지(H107), 4 정류부 정지(H103), 5 인버터 정지(H105, ESD 또는 절체 확인 뒤)
   - 먼저 확인해서 이미 그 상태면 명령하지 않는다. 명령 → i_tResend 기다림 → 안 됐으면 다시. 될 때까지 계속
   - i_tFail 넘게 안 되면 q_wFailed(오류)를 켠다. 오류가 켜져도 계속 보낸다. 되면 오류는 꺼진다
   - 드라이버가 못 받은 명령(바쁨·통신 끊김)은 기다리지 않고 다음 스캔에 다시 보낸다 (보낸 횟수에 넣지 않음)
   - 된 동작은 원인이 사라졌다가 다시 생길 때까지 다시 하지 않는다 (사람이 다시 켠 것을 되돌리지 않음)
   - UPS 명령은 스캔마다 하나. 순서는 바이패스 → 인버터(절체 확인 뒤) → BBC → 정류부: 앞 동작이 되거나 오류가 켜져야 다음 동작을 보낸다
     BMS는 전부 열기가 필요하면 충전만 열기는 하지 않는다
   - ESD나 화재가 걸려 있으면: 바이패스 절체는 하지 않는다(다른 원인이 요구해도). UPS 명령은 앞 동작을 기다리지 않고
     인버터 → BBC → 정류부 순으로 연달아 보낸다
   - i_bEnable(전체 스위치 AND 쓰기 관문)이 꺼지면 모두 처음 상태로
   - UPS 명령은 i_ipUps로 직접 보낸다. BMS 명령은 q_eBmsReq(그 스캔만)로 내고 MAIN이 드라이버를 부른다
   - 복귀(다시 켜기), MCCB Trip, 바이패스 포함 출력 차단, BMS E-stop은 하지 않는다
   변경: 2026-11-25 이중화 절체 때 상대의 된 동작 기억을 이어받음 (명세 RED-01·SQ-05 v2.49): i_bInheritLoad 때 i_wInheritDone을 담아 두고,
         그 동작이 필요해지면 보내지 않고 '됨'으로 둠 (사람이 다시 켠 것을 되돌리지 않음). 쓰기 허가·UPS 읽기 뒤 i_tInheritSettle 동안 안 쓰인 비트와
         i_tInheritMax가 지난 비트는 버림 *)
VAR_INPUT
	i_bEnable		: BOOL;					// GVL_PERSIST.g_bUpsSafetyRespEnable AND 장비 쓰기 관문
	i_nCause		: UDINT;				// FB_UpsSafetyStage.q_nRespCause (대응 원인, v2.30)
	i_stUps			: ST_UpsPublish_V1;		// UPS 보고값 (RectStatus b0, BBCStatus b0, InverterStatus b0, BypassStatus b0)
	i_bUpsValid		: BOOL;					// UPS 통신 정상
	i_stBms			: ST_EsolutionState;	// BMS 상태 (컨택터 30026·30027)
	i_ipUps			: I_Ups;				// UPS 명령 대상
	i_tResend		: TIME := T#2S;			// 보낸 뒤 다시 보내기까지 (응답 대기 1초 + 쉼 1초)
	i_tFail			: TIME := T#10S;		// 이 시간 넘게 안 되면 오류 표시 (보내기는 계속)
	i_bInheritLoad	: BOOL;					// 이 스캔에 이어받을 기억을 담음 (이중화: 이 PLC가 Active가 되는 순간, 명세 RED-01 v2.49)
	i_wInheritDone	: WORD;					// 이어받을 된 동작 비트 (대기 중 받은 상대의 q_wDone)
	i_tInheritSettle: TIME := T#3S;			// 쓰기 허가 + UPS 읽기 뒤 이 시간 동안 필요해지지 않은 이어받은 비트는 버림
	i_tInheritMax	: TIME := T#30S;		// 이어받은 비트는 담은 뒤 이 시간이 지나면 버림
END_VAR
VAR_OUTPUT
	q_wNeeded		: WORD;					// 지금 필요한 동작 (비트 0~5)
	q_wDone			: WORD;					// 된 동작
	q_wFailed		: WORD;					// 오류: i_tFail 넘게 안 된 동작 (계속 보내는 중. EMS 칸 없음, PLC 안에서만)
	q_eBmsReq		: UINT;					// BMS 요청: 0 없음, 1 충전 컨택터 열기, 2 전부 열기 (MAIN이 드라이버에 전달)
	q_nBmsSeq		: UDINT;				// 전부 열기 명령 번호 (M_SetStateCmd 중복 거르기용, 16#7F000000부터)
	q_anTry			: ARRAY[0..5] OF UINT;	// 동작별 보낸 횟수 (드라이버가 받은 것만, 65535에서 멈춤)
	q_bEsd			: BOOL;					// ESD·화재 대응 중 (순서 기다리지 않음, 바이패스 절체 안 함, v2.31 화재 포함)
	q_bBypassBlocked : BOOL;				// 바이패스 이상이라 바이패스 절체를 보내지 않는 중 (기록 BypassBlocked, v2.31)
	q_wInherit		: WORD;					// 아직 쓰지 않은 이어받은 된 동작 비트 (v2.49)
END_VAR
VAR
	_anState		: ARRAY[0..5] OF UINT;	// 0 보낼 차례, 1 보낸 뒤 기다림, 2 됨
	_atonResend		: ARRAY[0..5] OF TON;
	_atonFail		: ARRAY[0..5] OF TON;
	_abAchieved		: ARRAY[0..5] OF BOOL;
	_k				: INT;
	_i				: INT;
	_bNeed			: BOOL;
	_bUpsSent		: BOOL;					// 이번 스캔에 UPS 명령을 이미 시도함
	_bUpsHold		: BOOL;					// 앞 UPS 동작이 진행 중이라 뒤 동작은 기다림 (ESD가 아닐 때)
	_nBmsCount		: UDINT;
	_wBit			: WORD;
	_eCmd			: E_UpsCommand;
	_bInvStopArmed	: BOOL;					// 인버터 정지 To Bypass: 바이패스가 확인돼 인버터 정지를 시작함 (원인이 사라질 때까지 유지)
	_wInherit		: WORD;					// 이어받은 된 동작 비트 (쓰거나 버리면 지움, v2.49)
	_tonInheritSettle : TON;
	_tonInheritMax	: TON;
END_VAR
VAR CONSTANT
	ACT_CHG_OPEN	: INT := 0;
	ACT_BMS_OPEN	: INT := 1;
	ACT_BYPASS		: INT := 2;
	ACT_BBC_OFF		: INT := 3;
	ACT_RECT_OFF	: INT := 4;
	ACT_INV_OFF		: INT := 5;
	// 진행 순서 (동작 번호). UPS는 바이패스 → 인버터 → BBC → 정류부
	ORDER			: ARRAY[0..5] OF INT := [0, 1, 2, 5, 3, 4];
	// SQ-01 원인 비트
	C_BMS_MINOR		: UDINT := 16#00000004;	// b2
	C_BBC_GROUP		: UDINT := 16#00000388;	// b3 BMS Major, b7 지락(RCD)1, b8 BBC 중고장, b9 지락(RCD)2
	C_RECT			: UDINT := 16#00000010;	// b4 입력·정류부 중고장
	C_INV			: UDINT := 16#00002060;	// b5 출력, b6 인버터 중고장, b13 MBS C/B Fail → 바이패스 절체
	C_INV_STOP		: UDINT := 16#00002460;	// b5, b6, b13 MBS: 맵 '인버터정지 To Bypass', b10 BMS Level 3: 7쪽 표 5단계 '인버터 정지/바이패스 절체' (v2.54) → 절체 확인 뒤 인버터 정지 (화재는 v2.31부터 ESD처럼)
	C_FULL			: UDINT := 16#00000400;	// b10 BMS Level 3 (화재는 v2.31부터 C_ESD)
	C_ESD			: UDINT := 16#00001800;	// b11 화재, b12 ESD: 바이패스 절체 안 함, 인버터·BBC·정류부 정지 + BMS 전부 열기 (v2.31)
	W1_BYPASS		: UDINT := 16#03FF0000;	// UPS Warning1 b16~25 = I49 바이패스 이상 (맵 'To Bypass 절체 안 됨')
	BMS_SEQ_BASE	: UDINT := 16#7F000000;
END_VAR

// 이중화 이어받기 (명세 RED-01·SQ-05 v2.49): 담고, 오래되면 버림
IF i_bInheritLoad THEN
	_wInherit := i_wInheritDone AND 16#003F;
	_tonInheritSettle(IN := FALSE);
	_tonInheritMax(IN := FALSE);
END_IF
_tonInheritSettle(IN := _wInherit <> 0 AND i_bEnable AND i_bUpsValid, PT := i_tInheritSettle);
_tonInheritMax(IN := _wInherit <> 0, PT := i_tInheritMax);
IF _tonInheritSettle.Q OR _tonInheritMax.Q THEN
	_wInherit := 0;
END_IF

// 0) 됐는지 (확인 신호를 믿을 수 없으면 안 된 것으로 봄)
_abAchieved[ACT_CHG_OPEN] := i_stBms.bContactorFeedbackKnown AND NOT i_stBms.bChargeContactorClosed;
_abAchieved[ACT_BMS_OPEN] := i_stBms.bContactorFeedbackKnown AND i_stBms.wSystemContactor = 0 AND i_stBms.wRackContactor = 0;
_abAchieved[ACT_BYPASS] := i_bUpsValid AND i_stUps.BypassStatus.0;
_abAchieved[ACT_BBC_OFF] := i_bUpsValid AND NOT i_stUps.BBCStatus.0;
_abAchieved[ACT_RECT_OFF] := i_bUpsValid AND NOT i_stUps.RectStatus.0;
_abAchieved[ACT_INV_OFF] := i_bUpsValid AND NOT i_stUps.InverterStatus.0;

// 1) 원인 → 필요한 동작
q_wNeeded := 0;
q_bBypassBlocked := FALSE;
q_bEsd := i_bEnable AND (i_nCause AND C_ESD) <> 0;
IF i_bEnable THEN
	IF (i_nCause AND C_BMS_MINOR) <> 0 THEN q_wNeeded := q_wNeeded OR SHL(WORD#1, ACT_CHG_OPEN); END_IF
	IF (i_nCause AND C_BBC_GROUP) <> 0 THEN q_wNeeded := q_wNeeded OR SHL(WORD#1, ACT_BBC_OFF); END_IF
	IF (i_nCause AND C_RECT) <> 0 THEN
		q_wNeeded := q_wNeeded OR SHL(WORD#1, ACT_RECT_OFF) OR SHL(WORD#1, ACT_CHG_OPEN);
	END_IF
	IF (i_nCause AND C_INV) <> 0 THEN q_wNeeded := q_wNeeded OR SHL(WORD#1, ACT_BYPASS); END_IF
	IF (i_nCause AND C_FULL) <> 0 THEN
		q_wNeeded := q_wNeeded OR SHL(WORD#1, ACT_BYPASS) OR SHL(WORD#1, ACT_BBC_OFF) OR SHL(WORD#1, ACT_RECT_OFF) OR SHL(WORD#1, ACT_BMS_OPEN);
	END_IF
	// 인버터 정지 To Bypass (v2.30): 바이패스가 확인된 뒤에만 시작. 시작하면 원인이 사라질 때까지 유지
	IF (i_nCause AND C_INV_STOP) = 0 THEN
		_bInvStopArmed := FALSE;
	ELSIF _abAchieved[ACT_BYPASS] OR (_wInherit AND SHL(WORD#1, ACT_INV_OFF)) <> 0 THEN	// v2.49: 인버터 정지를 이어받으면 바이패스 확인을 기다리지 않음
		_bInvStopArmed := TRUE;
	END_IF
	IF _bInvStopArmed THEN q_wNeeded := q_wNeeded OR SHL(WORD#1, ACT_INV_OFF); END_IF
	// 바이패스 이상 (v2.31, O-17): 아직 바이패스가 아니면 절체를 보내지 않음 (부하는 인버터로 유지). 바이패스가 정상이 되면 다시 필요해짐
	IF NOT q_bEsd AND (q_wNeeded AND SHL(WORD#1, ACT_BYPASS)) <> 0 AND NOT _abAchieved[ACT_BYPASS]
		AND i_bUpsValid AND (i_stUps.Warning1 AND W1_BYPASS) <> 0 THEN
		q_bBypassBlocked := TRUE;
		q_wNeeded := q_wNeeded AND NOT SHL(WORD#1, ACT_BYPASS);
	END_IF
	IF q_bEsd THEN
		q_wNeeded := q_wNeeded OR SHL(WORD#1, ACT_INV_OFF) OR SHL(WORD#1, ACT_BBC_OFF) OR SHL(WORD#1, ACT_RECT_OFF) OR SHL(WORD#1, ACT_BMS_OPEN);
		q_wNeeded := q_wNeeded AND NOT SHL(WORD#1, ACT_BYPASS);	// 비상정지 중에 부하를 바이패스로 다시 살리지 않음
	END_IF
	IF (q_wNeeded AND SHL(WORD#1, ACT_BMS_OPEN)) <> 0 THEN
		q_wNeeded := q_wNeeded AND NOT SHL(WORD#1, ACT_CHG_OPEN);	// 전부 열기가 충전 열기를 포함
	END_IF
ELSE
	_bInvStopArmed := FALSE;
END_IF

// 2) 동작별 진행 (ORDER 순서)
_bUpsSent := FALSE;
_bUpsHold := FALSE;
q_eBmsReq := 0;
FOR _k := 0 TO 5 DO
	_i := ORDER[_k];
	_wBit := SHL(WORD#1, _i);
	_bNeed := (q_wNeeded AND _wBit) <> 0;
	_atonResend[_i](IN := _bNeed AND _anState[_i] = 1, PT := i_tResend);
	IF NOT _bNeed THEN
		_anState[_i] := 0;		// 원인이 사라짐 (또는 꺼짐) → 다음에 다시 생기면 처음부터
		q_anTry[_i] := 0;
	ELSE
		CASE _anState[_i] OF
			0:	// 보낼 차례
				IF (_wInherit AND _wBit) <> 0 THEN
					_anState[_i] := 2;	// 상대가 이미 한 동작 (이중화 이어받기, v2.49): 다시 보내지 않음
					_wInherit := _wInherit AND NOT _wBit;
				ELSIF _abAchieved[_i] THEN
					_anState[_i] := 2;	// 이미 그 상태
				ELSIF _i = ACT_CHG_OPEN OR _i = ACT_BMS_OPEN THEN
					IF q_eBmsReq = 0 THEN
						IF _i = ACT_BMS_OPEN THEN
							q_eBmsReq := 2;
							_nBmsCount := _nBmsCount + 1;
							q_nBmsSeq := BMS_SEQ_BASE + (_nBmsCount AND 16#00FFFFFF);
						ELSE
							q_eBmsReq := 1;
						END_IF
						IF q_anTry[_i] < 65535 THEN q_anTry[_i] := q_anTry[_i] + 1; END_IF
						_anState[_i] := 1;
					END_IF
				ELSIF NOT _bUpsSent AND NOT _bUpsHold AND i_ipUps <> 0 THEN
					CASE _i OF
						ACT_BYPASS:		_eCmd := E_UpsCommand.ToBypass;
						ACT_BBC_OFF:	_eCmd := E_UpsCommand.BbcOff;
						ACT_RECT_OFF:	_eCmd := E_UpsCommand.RectifierOff;
						ACT_INV_OFF:	_eCmd := E_UpsCommand.InverterOff;
					END_CASE
					_bUpsSent := TRUE;	// UPS는 스캔마다 하나
					IF i_ipUps.M_RequestCommand(_eCmd) THEN
						IF q_anTry[_i] < 65535 THEN q_anTry[_i] := q_anTry[_i] + 1; END_IF
						_anState[_i] := 1;
					END_IF	// 못 받았으면 0에 남아 다음 스캔에 다시
				END_IF
			1:	// 보낸 뒤 기다림
				IF _abAchieved[_i] THEN
					_anState[_i] := 2;
				ELSIF _atonResend[_i].Q THEN
					_anState[_i] := 0;	// 다시 보냄
				END_IF
		END_CASE
	END_IF
	_atonFail[_i](IN := _bNeed AND _anState[_i] <> 2, PT := i_tFail);
	// ESD가 아니면 앞 UPS 동작이 되거나 오류가 켜질 때까지 뒤 UPS 동작은 기다림
	IF _i >= ACT_BYPASS AND _bNeed AND _anState[_i] <> 2 AND NOT _atonFail[_i].Q AND NOT q_bEsd THEN
		_bUpsHold := TRUE;
	END_IF
END_FOR

q_wDone := 0;
q_wFailed := 0;
FOR _i := 0 TO 5 DO
	IF _anState[_i] = 2 THEN q_wDone := q_wDone OR SHL(WORD#1, _i); END_IF
	IF _atonFail[_i].Q THEN q_wFailed := q_wFailed OR SHL(WORD#1, _i); END_IF
END_FOR
q_wInherit := _wInherit;

END_FUNCTION_BLOCK

// ---- 20_Module/Ups/FB_UpsSafetyStage.TcPOU
(* LiB-UPS 사고·고장 단계 판정 (④보호 표시 / 장치: UPS·BAT). 2026-11-05.
   기반 없음(신규). 동작시퀀스 7쪽(이솔루션 2026-10-23) 단계표를 따른다.
   변경: 2026-11-09 UPS 경고·고장 4번 칸을 없앰. STATUS 비트를 Warning3 하위·Fault3 상위에서 읽음 (명세 RD-UPS-02 v1.6)
   변경: 2026-11-18 UPS 경고·고장 칸을 회사 eventMap 순서로 읽음 (Warning1·Fault1·Fault2, 명세 RD-UPS-02 v2.20)
   변경: 2026-11-18 기록(FB_UpsSafetyLog)용 출력 q_nLatched·q_bAckPulse·q_nAckCleared 추가 (명세 SQ-01 v2.21). 판정은 그대로
   변경: 2026-11-20 대응(SQ-05)용 원인 q_nRespCause 추가 (명세 SQ-05 v2.30, 세방 맵 Alarm Flag 비트별 동작). 단계 판정은 그대로
         - b4: '기동 안 됨' 2비트(Fault1 b7 입력 상회전, b18 Pre Magnet Fail) 뺌
         - b5: 출력 과전류 R/S/T(Fault2 b0~2)는 i_tOutOcDelay(15분) 계속될 때만, 출력 과전류 Trip(b3~5)은 바로
         - b8: 배터리 과전류(Fault1 b23)는 i_tBattOcDelay(10분) 계속될 때만, 나머지 BBC 중고장은 바로
         - b13: MBS C/B Fail(Fault2 b14, I50 b7). 단계 없음, 대응만
   변경: 2026-11-23 Fault(4~6단계)도 원인이 풀리면 바로 내림. 확인 전 유지(래치)와 i_bAck·q_bAckPending·q_nLatched·q_bAckPulse·q_nAckCleared 없앰
         (명세 SQ-01 v2.38: 확인은 EMS가 하므로 PMS에 확인 신호가 오지 않아, 붙잡은 Fault가 재시작 전까지 안 풀렸음)
   변경: 2026-11-23 i_bClear 추가: 이중화 대기 중에는 원인을 비움 (명세 RED-02 v2.45: 장비를 읽지 않으니 마지막 값이 옛 값. 넘겨받는 순간 옛 값으로 대응하지 않게)
   부호·단위: 해당 없음. 명세: C:\gil\UPS\명세작업\UPS_명세서.md SQ-01, SQ-05
   차단·정지는 UPS(UMS)와 BMS가 스스로 한다. 이 FB는 판정과 표시만 하고 장비에 아무것도 쓰지 않는다. *)
FUNCTION_BLOCK FB_UpsSafetyStage
VAR_INPUT
	i_stUps			: ST_UpsPublish_V1;	// UPS 보고값 (FB_RptSebangUps.q_stUps)
	i_bUpsValid		: BOOL;				// UPS 데이터 유효 (통신 정상)
	i_stBat			: ST_BatPublish_V1;	// 짝 BAT 보고값 (FB_RptEsolutionBat.q_stBat)
	i_bBatValid		: BOOL;				// BAT 데이터 유효 (통신 정상)
	i_tOutOcDelay	: TIME := T#15M;	// 출력 과전류 R/S/T가 이만큼 계속되면 대응 (세방 맵 '15분후 인버터정지 To Bypass', SQ-05 v2.30)
	i_bClear		: BOOL;				// 원인을 비움 (이중화 대기 중, 명세 RED-02 v2.45). 통신 끊김 때 마지막 값 유지보다 우선
	i_tBattOcDelay	: TIME := T#10M;	// 배터리 과전류가 이만큼 계속되면 대응 (세방 맵 '10분후 정지', SQ-05 v2.30)
END_VAR
VAR_OUTPUT
	q_nStage		: UINT;				// 대표 단계 0~6 (걸린 단계 중 가장 높은 것)
	q_wStageMask	: WORD;				// 걸린 단계 목록. bit n = n단계 (n = 1~6). 높은 순서로 모두 표시할 때 사용
	q_nCause		: UDINT;			// 원인 비트 (아래 CAUSE_* 표). q_nActiveCause와 같음 (v2.38: Fault도 붙잡지 않음)
	q_nActiveCause	: UDINT;			// 지금 실제로 걸린 원인만
	q_bUpsCommFault	: BOOL;				// UPS 통신장애 (단계와 별도 상태). 끊긴 동안 UPS 원인은 마지막 값을 유지
	q_bBatCommFault	: BOOL;				// BAT 통신장애 (단계와 별도 상태). 끊긴 동안 BAT 원인은 마지막 값을 유지
	q_nRespCause	: UDINT;			// 대응(FB_UpsSafetyResponse)용 원인. 비트 배치는 q_nActiveCause와 같고 b13 MBS C/B Fail 추가 (SQ-05 v2.30)
END_VAR
VAR
	_nUpsCause		: UDINT;			// UPS에서 나온 원인 (통신이 끊기면 마지막 값 유지)
	_nBatCause		: UDINT;			// BAT에서 나온 원인 (통신이 끊기면 마지막 값 유지)
	_nUpsResp		: UDINT;			// UPS에서 나온 대응 원인 (통신이 끊기면 마지막 값 유지)
	_tonOutOc		: TON;				// 출력 과전류 R/S/T 지속
	_tonBattOc		: TON;				// 배터리 과전류 지속
	_i				: INT;
END_VAR
VAR CONSTANT
	(* 원인 비트 → 단계. 순서 = 비트 번호 *)
	CAUSE_STAGE		: ARRAY[0..12] OF UINT := [
		1,	// b0  AC·DC SPD (I51 b8·b9)
		1,	// b1  UPS 경고장 (SPD·BMS Minor 제외)
		2,	// b2  BMS Minor (I51 b10)
		3,	// b3  BMS Major (I51 b11)
		3,	// b4  UPS 입력·정류부 중고장 (I44·I45)
		3,	// b5  UPS 출력 중고장 (I47)
		3,	// b6  UPS 인버터 중고장 (I48)
		3,	// b7  배터리 DC 전로 지락(RCD) 1단계 (I51 b12, 명세 v2.50 세방 회신)
		4,	// b8  배터리 컨버터(BBC) 중고장 (I46)
		4,	// b9  배터리 DC 전로 지락(RCD) 2단계 (I51 b13, 명세 v2.50 세방 회신)
		5,	// b10 BMS Level 3 (BAT Status b9 System Lock)
		5,	// b11 화재 (I51 b14)
		6];	// b12 ESD (I50 b0)
	(* UPS 보고 칸 안의 비트 (명세 RD-UPS-02 v2.20, 회사 eventMap 순서) *)
	W1_SPD			: UDINT := 16#18000000;	// Warning1 b27 AC SPD (I51 b8), b28 DC SPD (I51 b9)
	W1_BMS_MINOR	: UDINT := 16#20000000;	// Warning1 b29 BMS Minor (I51 b10)
	F1_INPUT		: UDINT := 16#003FFFFF;	// Fault1 b0~b21 입력·정류부 (I44·I45)
	F1_BBC			: UDINT := 16#3FC00000;	// Fault1 b22~b29 배터리 컨버터 (I46)
	F2_OUTPUT		: UDINT := 16#0000003F;	// Fault2 b0~b5 출력 (I47)
	F2_INVERTER		: UDINT := 16#00001FC0;	// Fault2 b6~b12 인버터 (I48)
	F2_ESD			: UDINT := 16#00002000;	// Fault2 b13 Emergency Stop (I50 b0). b14 MBS C/B Fail (I50 b7)은 단계 없음
	F2_BMS_MAJOR	: UDINT := 16#00008000;	// Fault2 b15 BMS Major (I51 b11)
	F2_RCD1			: UDINT := 16#00010000;	// Fault2 b16 지락(RCD) 1단계 (I51 b12)
	F2_RCD2			: UDINT := 16#00020000;	// Fault2 b17 지락(RCD) 2단계 (I51 b13)
	F2_FIRE			: UDINT := 16#00040000;	// Fault2 b18 화재 (I51 b14)
	(* 대응 원인 (SQ-05 v2.30, 세방 맵 Alarm Flag 정류부·배터리컨버터·인버터 칸) *)
	F1_START_BLOCK	: UDINT := 16#00040080;	// Fault1 b7 입력 상회전 (I44 b7), b18 Pre Magnet Fail (I45 b9): 맵 '기동 안 됨' → 명령 없음
	F1_BATT_OC		: UDINT := 16#00800000;	// Fault1 b23 배터리 과전류 (I46 b4): 맵 '10분후 정지'
	F2_OUT_OC		: UDINT := 16#00000007;	// Fault2 b0~2 출력 과전류 R/S/T (I47 b8~10): 맵 '15분후 인버터정지 To Bypass'
	F2_MBS			: UDINT := 16#00004000;	// Fault2 b14 MBS C/B Fail (I50 b7): 맵 '인버터정지 To Bypass', 단계 없음
	RESP_MBS		: UDINT := 16#00002000;	// 대응 원인 b13 MBS C/B Fail
END_VAR

// 1) UPS 원인. 통신이 끊기면 마지막 값을 그대로 둔다 (단계를 내리지 않음)
q_bUpsCommFault := NOT i_bUpsValid;
IF i_bUpsValid THEN
	_nUpsCause := 0;
	IF (i_stUps.Warning1 AND W1_SPD) <> 0 THEN _nUpsCause := _nUpsCause OR 16#0001; END_IF
	IF ((i_stUps.Warning1 AND NOT (W1_SPD OR W1_BMS_MINOR)) OR i_stUps.Warning2 OR i_stUps.Warning3) <> 0 THEN _nUpsCause := _nUpsCause OR 16#0002; END_IF
	IF (i_stUps.Warning1 AND W1_BMS_MINOR) <> 0 THEN _nUpsCause := _nUpsCause OR 16#0004; END_IF
	IF (i_stUps.Fault2 AND F2_BMS_MAJOR) <> 0 THEN _nUpsCause := _nUpsCause OR 16#0008; END_IF
	IF (i_stUps.Fault1 AND F1_INPUT) <> 0 THEN _nUpsCause := _nUpsCause OR 16#0010; END_IF
	IF (i_stUps.Fault2 AND F2_OUTPUT) <> 0 THEN _nUpsCause := _nUpsCause OR 16#0020; END_IF
	IF (i_stUps.Fault2 AND F2_INVERTER) <> 0 THEN _nUpsCause := _nUpsCause OR 16#0040; END_IF
	IF (i_stUps.Fault2 AND F2_RCD1) <> 0 THEN _nUpsCause := _nUpsCause OR 16#0080; END_IF
	IF (i_stUps.Fault1 AND F1_BBC) <> 0 THEN _nUpsCause := _nUpsCause OR 16#0100; END_IF
	IF (i_stUps.Fault2 AND F2_RCD2) <> 0 THEN _nUpsCause := _nUpsCause OR 16#0200; END_IF
	IF (i_stUps.Fault2 AND F2_FIRE) <> 0 THEN _nUpsCause := _nUpsCause OR 16#0800; END_IF
	IF (i_stUps.Fault2 AND F2_ESD) <> 0 THEN _nUpsCause := _nUpsCause OR 16#1000; END_IF
	// 대응 원인 (SQ-05 v2.30): 단계 원인에서 b4·b5·b8을 맵 동작 기준으로 다시 정하고 b13을 더함
	_tonOutOc(IN := (i_stUps.Fault2 AND F2_OUT_OC) <> 0, PT := i_tOutOcDelay);
	_tonBattOc(IN := (i_stUps.Fault1 AND F1_BATT_OC) <> 0, PT := i_tBattOcDelay);
	_nUpsResp := _nUpsCause AND NOT UDINT#16#00000130;
	IF (i_stUps.Fault1 AND F1_INPUT AND NOT F1_START_BLOCK) <> 0 THEN _nUpsResp := _nUpsResp OR 16#0010; END_IF
	IF (i_stUps.Fault2 AND F2_OUTPUT AND NOT F2_OUT_OC) <> 0 OR _tonOutOc.Q THEN _nUpsResp := _nUpsResp OR 16#0020; END_IF
	IF (i_stUps.Fault1 AND F1_BBC AND NOT F1_BATT_OC) <> 0 OR _tonBattOc.Q THEN _nUpsResp := _nUpsResp OR 16#0100; END_IF
	IF (i_stUps.Fault2 AND F2_MBS) <> 0 THEN _nUpsResp := _nUpsResp OR RESP_MBS; END_IF
END_IF

// 2) BAT 원인
q_bBatCommFault := NOT i_bBatValid;
IF i_bBatValid THEN
	_nBatCause := 0;
	IF i_stBat.Status.9 THEN _nBatCause := _nBatCause OR 16#0400; END_IF	// BMS Level 3 (System Lock)
END_IF

// 이중화 대기 중: 원인과 지연 타이머를 비움 (명세 RED-02 v2.45)
IF i_bClear THEN
	_nUpsCause := 0;
	_nBatCause := 0;
	_nUpsResp := 0;
	_tonOutOc(IN := FALSE, PT := i_tOutOcDelay);
	_tonBattOc(IN := FALSE, PT := i_tBattOcDelay);
END_IF
q_nActiveCause := _nUpsCause OR _nBatCause;
q_nRespCause := _nUpsResp OR _nBatCause;

// 3) Warning·Fault 모두 원인이 풀리면 바로 내림 (v2.38. 확인은 EMS가 함). 통신이 끊긴 장비 원인은 위에서 마지막 값 유지
q_nCause := q_nActiveCause;

// 4) 단계 목록과 대표 단계
q_wStageMask := 0;
q_nStage := 0;
FOR _i := 0 TO 12 DO
	IF (q_nCause AND SHL(UDINT#1, _i)) <> 0 THEN
		q_wStageMask := q_wStageMask OR SHL(WORD#1, CAUSE_STAGE[_i]);
		q_nStage := MAX(q_nStage, CAUSE_STAGE[_i]);
	END_IF
END_FOR

END_FUNCTION_BLOCK

// ---- 20_Module/Ups/FB_UpsSafetyLog.TcPOU
FUNCTION_BLOCK FB_UpsSafetyLog		// UPS 사고·고장 단계 기록: FB_UpsSafetyStage 결과를 PMS 이벤트 로그에 남김 (EMS로는 안 보냄)
(* 사고·고장 단계·원인 기록 (④보호 표시 / 장치: UPS·BAT). 2026-11-18.
   기반: 예전 작업본 pms-standard-main FB_UpsSafetyLog (2026-11-09, 명세 v2.0). 저장소 밖 C:\gil\UPS_보관\pms-standard-main
   변경: UPSstd로 옮김. 기록은 PMS 이벤트 로그(TwinCAT 이벤트 로거, XAE Error List)에만. 이벤트 클래스 PmsUps는
     로거 리스너(FB_MqttLoggerListener)가 받지 않아 EMS(pms_log)로 가지 않는다 (명세 SQ-01 v2.21).
     시험용 출력 q_bSettled 등과 안정 시간 입력 i_tSettle을 더함.
   변경: 2026-11-19 대응 동작(FB_UpsSafetyResponse) 기록 추가: 처음 보낸 명령, 완료, 10초 오류 (명세 SQ-01·SQ-05 v2.22)
   변경: 2026-11-23 확인 대기(AckPending)·Fault 확인(FaultAck) 기록 없앰. PMS 안에서 Fault를 붙잡지 않음 (명세 SQ-01 v2.38)
   부호·단위: 해당 없음. 명세: C:\gil\UPS\명세작업\UPS_명세서.md SQ-01 "기록"
   - 원인 알람(CauseActive): 원인 비트마다 발생·해소 1회 ("UPS n 사고·고장 k단계: 원인"). 심각도 1~3단계 Warning, 4~5 Error, 6 Critical
   - 단계 바뀜(StageChange): 대표 단계가 바뀔 때마다 메시지 1회
   - 통신장애(CommLost): 한 번이라도 통신이 됐던 장비가 끊겼을 때만 알람 (설치 안 된 장비는 기록 안 함)
   - 대응 명령(RespCmd): 동작을 처음 보낼 때 1번. 2초마다 다시 보내는 것은 남기지 않음 (보낸 횟수 0 → 1 이상)
   - 대응 완료(RespDone): 동작이 될 때 1번 (보낸 횟수, 보내기 전에 이미 그 상태였으면 그렇게)
   - 대응 오류(RespFail): 10초 넘게 안 된 동작마다 알람. 되거나 필요 없어지면 해소
   - 바이패스 절체 안 함(BypassBlocked): 바이패스 이상이라 절체를 보내지 않는 동안 알람 (명세 SQ-05 v2.31, 2026-11-20)
   - 켜진 뒤 i_tSettle 동안은 기록하지 않음 (부팅 직후 통신이 붙기 전 값으로 기록하지 않기 위해)
   판정은 하지 않는다. 원인 비트 순서·단계는 FB_UpsSafetyStage.CAUSE_STAGE와 같아야 한다 *)
VAR_INPUT
	i_nUps			: UINT;					// UPS 번호 (1~)
	i_nStage		: UINT;					// FB_UpsSafetyStage.q_nStage
	i_nActiveCause	: UDINT;				// FB_UpsSafetyStage.q_nActiveCause
	i_bUpsCommFault	: BOOL;					// FB_UpsSafetyStage.q_bUpsCommFault
	i_bBatCommFault	: BOOL;					// FB_UpsSafetyStage.q_bBatCommFault
	i_wRespNeeded	: WORD;					// FB_UpsSafetyResponse.q_wNeeded (지금 필요한 동작, 비트 0~5)
	i_wRespDone		: WORD;					// FB_UpsSafetyResponse.q_wDone
	i_wRespFailed	: WORD;					// FB_UpsSafetyResponse.q_wFailed (10초 넘게 안 된 동작)
	i_anRespTry		: ARRAY[0..5] OF UINT;	// FB_UpsSafetyResponse.q_anTry (동작별 보낸 횟수)
	i_bBypassBlocked : BOOL;				// FB_UpsSafetyResponse.q_bBypassBlocked (v2.31)
	i_tSettle		: TIME := T#15S;		// 켜진 뒤 기록하지 않는 시간
END_VAR
VAR_OUTPUT
	q_bSettled		: BOOL;					// 기록 시작함 (i_tSettle 지남)
	q_nRaised		: UDINT;				// 원인 알람이 발생 중인 원인 비트
	q_bUpsCommRaised : BOOL;				// UPS 통신장애 알람 발생 중
	q_bBatCommRaised : BOOL;				// BMS 통신장애 알람 발생 중
	q_nStageMsg		: UDINT;				// 단계 바뀜 메시지 보낸 수
	q_nRespCmdMsg	: UDINT;				// 대응 명령 메시지 보낸 수
	q_nRespDoneMsg	: UDINT;				// 대응 완료 메시지 보낸 수
	q_wRespFailRaised : WORD;				// 대응 오류 알람이 발생 중인 동작 비트
	q_bBypassBlockedRaised : BOOL;			// 바이패스 절체 안 함 알람 발생 중
END_VAR
VAR
	_tonSettle		: TON;
	_afbCause		: ARRAY[0..12] OF FB_LogAlarm;
	_fbUpsComm		: FB_LogAlarm;
	_fbBatComm		: FB_LogAlarm;
	_fbStage		: FB_LogMsg;
	_bUpsEverOk		: BOOL;
	_bBatEverOk		: BOOL;
	_nLastStage		: UINT;
	_asArg			: ARRAY[1..6] OF WSTRING(63);
	_stEntry		: TcEventEntry;
	_i				: INT;
	_bActive		: BOOL;
	_afbRespFail	: ARRAY[0..5] OF FB_LogAlarm;
	_fbRespCmd		: FB_LogMsg;
	_fbRespDone		: FB_LogMsg;
	_fbBypassBlocked : FB_LogAlarm;
	_wSent			: WORD;					// 한 번이라도 보낸 동작 (보낸 횟수 > 0)
	_wSentLast		: WORD;
	_wDone			: WORD;					// 필요하고 된 동작
	_wDoneLast		: WORD;
	_wBit			: WORD;
END_VAR
VAR CONSTANT
	CAUSE_STAGE		: ARRAY[0..12] OF UINT := [1, 1, 2, 3, 3, 3, 3, 3, 4, 4, 5, 5, 6];	// FB_UpsSafetyStage와 같음
	CAUSE_NAME		: ARRAY[0..12] OF WSTRING(31) := [
		"SPD", "UPS 경고장", "BMS Minor", "BMS Major", "입력·정류부 중고장", "출력 중고장", "인버터 중고장",
		"지락(RCD) 1단계", "배터리 컨버터 중고장", "지락(RCD) 2단계", "BMS Level 3", "화재", "ESD"];
	(* 대응 동작 이름 = FB_UpsSafetyResponse 동작 번호 순서 (명세 SQ-05) *)
	RESP_NAME		: ARRAY[0..5] OF WSTRING(39) := [
		"충전 컨택터 열기(BMS 40014=0)", "BMS 컨택터 전부 열기(40013~15=0)", "바이패스 절체(H109)",
		"BBC 정지(H107)", "정류부 정지(H103)", "인버터 정지(H105)"];
END_VAR

IF NOT i_bUpsCommFault THEN _bUpsEverOk := TRUE; END_IF
IF NOT i_bBatCommFault THEN _bBatEverOk := TRUE; END_IF
_tonSettle(IN := TRUE, PT := i_tSettle);
q_bSettled := _tonSettle.Q;
_wSent := 0;
FOR _i := 0 TO 5 DO
	IF i_anRespTry[_i] > 0 THEN _wSent := _wSent OR SHL(WORD#1, _i); END_IF
END_FOR
_wDone := i_wRespDone AND i_wRespNeeded;
IF NOT q_bSettled THEN
	_nLastStage := i_nStage;
	_wSentLast := _wSent;
	_wDoneLast := _wDone;
	RETURN;
END_IF

// 1) 원인 알람 (지금 실제로 걸린 원인)
q_nRaised := 0;
FOR _i := 0 TO 12 DO
	_bActive := (i_nActiveCause AND SHL(UDINT#1, _i)) <> 0;
	IF _bActive <> _afbCause[_i].q_bRaised THEN
		_asArg[1] := TO_WSTRING(i_nUps);
		_asArg[2] := TO_WSTRING(CAUSE_STAGE[_i]);
		_asArg[3] := CAUSE_NAME[_i];
	END_IF
	_stEntry := TC_EVENTS.PmsUps.CauseActive;
	IF CAUSE_STAGE[_i] >= 6 THEN
		_stEntry.eSeverity := TcEventSeverity.Critical;
	ELSIF CAUSE_STAGE[_i] >= 4 THEN
		_stEntry.eSeverity := TcEventSeverity.Error;
	ELSE
		_stEntry.eSeverity := TcEventSeverity.Warning;
	END_IF
	_afbCause[_i](i_stEntry := _stEntry, i_bActive := _bActive, i_nArgs := 3, i_asArg := _asArg);
	IF _afbCause[_i].q_bRaised THEN
		q_nRaised := q_nRaised OR SHL(UDINT#1, _i);
	END_IF
END_FOR

// 2) 대표 단계 바뀜
_fbStage(i_stEntry := TC_EVENTS.PmsUps.StageChange);
IF i_nStage <> _nLastStage THEN
	_asArg[1] := TO_WSTRING(i_nUps);
	_asArg[2] := TO_WSTRING(_nLastStage);
	_asArg[3] := TO_WSTRING(i_nStage);
	_fbStage.M_SendEvent(i_nArgs := 3, i_asArg := _asArg);
	_nLastStage := i_nStage;
	q_nStageMsg := q_nStageMsg + 1;
END_IF

// 3) 통신장애 (한 번이라도 됐던 장비만)
_bActive := i_bUpsCommFault AND _bUpsEverOk;
IF _bActive <> _fbUpsComm.q_bRaised THEN
	_asArg[1] := TO_WSTRING(i_nUps);
	_asArg[2] := "UPS";
END_IF
_fbUpsComm(i_stEntry := TC_EVENTS.PmsUps.CommLost, i_bActive := _bActive, i_nArgs := 2, i_asArg := _asArg);
q_bUpsCommRaised := _fbUpsComm.q_bRaised;
_bActive := i_bBatCommFault AND _bBatEverOk;
IF _bActive <> _fbBatComm.q_bRaised THEN
	_asArg[1] := TO_WSTRING(i_nUps);
	_asArg[2] := "BMS";
END_IF
_fbBatComm(i_stEntry := TC_EVENTS.PmsUps.CommLost, i_bActive := _bActive, i_nArgs := 2, i_asArg := _asArg);
q_bBatCommRaised := _fbBatComm.q_bRaised;

// 4) 대응 동작 (명세 SQ-05 기록, v2.22): 처음 보낸 명령, 완료, 10초 오류
_fbRespCmd(i_stEntry := TC_EVENTS.PmsUps.RespCmd);
_fbRespDone(i_stEntry := TC_EVENTS.PmsUps.RespDone);
q_wRespFailRaised := 0;
FOR _i := 0 TO 5 DO
	_wBit := SHL(WORD#1, _i);
	IF (_wSent AND _wBit) <> 0 AND (_wSentLast AND _wBit) = 0 THEN
		_asArg[1] := TO_WSTRING(i_nUps);
		_asArg[2] := RESP_NAME[_i];
		_fbRespCmd.M_SendEvent(i_nArgs := 2, i_asArg := _asArg);
		q_nRespCmdMsg := q_nRespCmdMsg + 1;
	END_IF
	IF (_wDone AND _wBit) <> 0 AND (_wDoneLast AND _wBit) = 0 THEN
		_asArg[1] := TO_WSTRING(i_nUps);
		_asArg[2] := RESP_NAME[_i];
		IF i_anRespTry[_i] = 0 THEN
			_asArg[3] := "이미 그 상태였음";
		ELSE
			_asArg[3] := WCONCAT("보낸 횟수 ", TO_WSTRING(i_anRespTry[_i]));
		END_IF
		_fbRespDone.M_SendEvent(i_nArgs := 3, i_asArg := _asArg);
		q_nRespDoneMsg := q_nRespDoneMsg + 1;
	END_IF
	_bActive := (i_wRespFailed AND _wBit) <> 0;
	IF _bActive <> _afbRespFail[_i].q_bRaised THEN
		_asArg[1] := TO_WSTRING(i_nUps);
		_asArg[2] := RESP_NAME[_i];
	END_IF
	_afbRespFail[_i](i_stEntry := TC_EVENTS.PmsUps.RespFail, i_bActive := _bActive, i_nArgs := 2, i_asArg := _asArg);
	IF _afbRespFail[_i].q_bRaised THEN
		q_wRespFailRaised := q_wRespFailRaised OR _wBit;
	END_IF
END_FOR
// 바이패스 이상이라 절체 안 함 (v2.31)
IF i_bBypassBlocked <> _fbBypassBlocked.q_bRaised THEN
	_asArg[1] := TO_WSTRING(i_nUps);
END_IF
_fbBypassBlocked(i_stEntry := TC_EVENTS.PmsUps.BypassBlocked, i_bActive := i_bBypassBlocked, i_nArgs := 1, i_asArg := _asArg);
q_bBypassBlockedRaised := _fbBypassBlocked.q_bRaised;
_wSentLast := _wSent;
_wDoneLast := _wDone;

END_FUNCTION_BLOCK

// ---- 20_Module/Mqtt/FB_EmsConfigApply.TcPOU
FUNCTION_BLOCK FB_EmsConfigApply		// EMS config(pcs·bat) → 운영 설정 (PlcTask. MAIN 액션 A_PassEmsCfg가 부름) [9-21 수정 2026-11-04: 추가]
(* - 입력 i_stCfg는 MAIN이 GVL_IF.g_stEmsCfg에서 일관되게 복사해 넘김. PCS·BMS 칸마다 번호(anPcsSeq·anBatSeq)가 바뀌면 새 레코드
   - [21번 수정 2026-11-09] is_available = 0인 값은 기본값으로 반영 (원래: 바꾸지 않고 기존 값 유지 → EMS가 한도를 풀 수 없었음)
       pcs 충전·방전 한도 0 → 그 방향 정격 (= 제한 없음). 두 방향 모두 0 → 그 PCS 유닛의 사용자 P 한도 끔 (bPEnable FALSE, 값은 ±정격)
       bat SOC 하한 0 → 0 %, 상한 0 → 100 % (감발 폭 fBand·재개 마진은 HMI 설정 그대로)
   - [UPS 2026-11-10] UPS 현장의 config/bat 레코드는 103.Config BAT UPS_V1 형식 (SocMin·SocMax = REAL, is_available 없음. UPS_MQTT_INTERFACE.md).
       그래서 bat 값은 받은 BMS(_abBatRx)만 계산에 넣고 항상 '있음'으로 봄. 아직 못 받은 BMS는 기본값(0 %·100 %)과 같아 결과에 영향 없음. pcs 쪽은 STD 그대로
   - pcs: 충전·방전 전력 한도 (kW) → 사용자 한도 stUnitLimit. 그 PCS의 유닛들에 정격 비율로 나눔, 충전은 fPMin (−). PvMarginRate는 쓰지 않음 (사양 대기)
   - bat: SOC 최소·최대 (%) → SOC 정책 stSocLimit. 배터리 그룹 전체 한 세트라 받은 BMS 값(기본값 포함) 중 가장 엄격한 값 (하한 = 가장 큰 값, 상한 = 가장 작은 값)
   - 범위 검사를 먼저 하고 통과한 값만 씀 (SOC는 FB_SocLimit.M_CheckSet과 같은 F_SocLimitSetErr). 버리면 q_bRejected (이벤트 로그 '잘못된 설정 값')
   - 쓴 값은 GVL_PERSIST라 재시작 뒤에도 남음. 설정 보호(FB_SettingGuard)가 한 번 더 지킴. 바꾸면 q_bApplied (이벤트 로그 '운영 설정 바뀜')
   - protection(배터리·배터리실 온도·습도 경고·고장)은 반영하지 않음 (값의 뜻·센서 대기. echo만)
   - M_BuildEcho: 설정 보호 뒤 실제 설정 → q_stEcho (MAIN이 GVL_IF.g_stEmsCfgEcho에 씀 → config echo) *)
VAR_INPUT
	i_bValid		: BOOL;			// 이번 스캔에 i_stCfg를 일관되게 복사함
	i_stCfg			: ST_IfEmsCfg;
	i_astUnitCfg	: ARRAY[1..GVL_PARAM.UNIT_COUNT] OF ST_UnitCfg;	// 유닛 ← PCS 번호, 정격
END_VAR
VAR_IN_OUT
	iq_stSocLimit	: ST_SocLimitSet;	// GVL_PERSIST.g_stModuleSet.stSocLimit
	iq_stUnitLimit	: ST_UnitLimitSet;	// GVL_PERSIST.g_stModuleSet.stUnitLimit
END_VAR
VAR_OUTPUT
	q_bApplied		: BOOL;			// 이번 스캔에 설정을 바꿈 (1스캔)
	q_sApplied		: WSTRING(63);
	q_bRejected		: BOOL;			// 이번 스캔에 받은 값을 버림 (1스캔)
	q_sRejected		: WSTRING(63);	// 마지막으로 버린 값과 이유
	q_nApplied		: UDINT;
	q_nRejected		: UDINT;
	q_stEcho		: ST_IfEmsCfgEcho;
END_VAR
VAR CONSTANT
	MAX_KW			: REAL := 1.0E6;	// kW. 이보다 큰 한도는 이상값
	SOC_MIN_DEFAULT	: REAL := 0.0;		// %, bat SocMin is_available 0일 때 [21번 수정 2026-11-09: 추가]
	SOC_MAX_DEFAULT	: REAL := 100.0;	// %, bat SocMax is_available 0일 때
END_VAR
VAR
	_stCfg			: ST_IfEmsCfg;		// 마지막으로 일관되게 받은 칸 (echo의 PvMarginRate)
	_anPcsSeq		: ARRAY[1..GVL_PARAM.PCS_COUNT] OF UDINT;
	_anBatSeq		: ARRAY[1..GVL_PARAM.BMS_COUNT] OF UDINT;
	_astBat			: ARRAY[1..GVL_PARAM.BMS_COUNT] OF ST_BatConfig_Rx;	// BMS마다 받아 둔 레코드 (가장 엄격한 SOC 계산)
	_astBatBefore	: ARRAY[1..GVL_PARAM.BMS_COUNT] OF ST_BatConfig_Rx;
	_abBatRx		: ARRAY[1..GVL_PARAM.BMS_COUNT] OF BOOL;	// [UPS] 그 BMS 레코드를 한 번이라도 받아 둠 (REAL 형식이라 빈 칸을 is_available로 못 가림)
	_abBatRxBefore	: ARRAY[1..GVL_PARAM.BMS_COUNT] OF BOOL;
	_stUnit			: ST_UnitLimitSet;
	_stSoc			: ST_SocLimitSet;
	_sErr			: WSTRING(63);
	p				: UINT;
	u				: UINT;
	b				: UINT;
	fSum			: REAL;
	fCh				: REAL;
	fDis			: REAL;
	fMin			: REAL;
	fMax			: REAL;
	bCh				: BOOL;
	bDis			: BOOL;
	bAny			: BOOL;
	bNewBat			: BOOL;
	bBad			: BOOL;
END_VAR

q_bApplied	:= FALSE;
q_bRejected	:= FALSE;
IF NOT i_bValid THEN
	RETURN;
END_IF
_stCfg := i_stCfg;

(* PCS: 충전·방전 전력 한도 → 그 PCS 유닛들의 사용자 한도 (정격 비율) *)
_stUnit := iq_stUnitLimit;
bAny := FALSE;
FOR p := 1 TO GVL_PARAM.PCS_COUNT DO
	IF i_stCfg.anPcsSeq[p] <> _anPcsSeq[p] THEN
		_anPcsSeq[p] := i_stCfg.anPcsSeq[p];
		bCh		:= i_stCfg.astPcs[p].ChargePowerLimit.is_available <> 0;
		bDis	:= i_stCfg.astPcs[p].DisChargePowerLimit.is_available <> 0;
		fCh		:= UDINT_TO_REAL(i_stCfg.astPcs[p].ChargePowerLimit.value);
		fDis	:= UDINT_TO_REAL(i_stCfg.astPcs[p].DisChargePowerLimit.value);
		fSum := 0.0;
		FOR u := 1 TO GVL_PARAM.UNIT_COUNT DO
			IF i_astUnitCfg[u].nPcs = p AND F_RealOk(i_astUnitCfg[u].fPRated) THEN
				fSum := fSum + i_astUnitCfg[u].fPRated;
			END_IF
		END_FOR
		IF (bCh AND fCh > MAX_KW) OR (bDis AND fDis > MAX_KW) THEN
			M_Reject(F_TxtNum("EMS config pcs 전력 한도 범위 밖: PCS ", p));
		ELSIF NOT (fSum > 0.0) THEN
			M_Reject(F_TxtNum("EMS config pcs 유닛 없음(정격 합 0): PCS ", p));
		ELSE
			// [21번 수정 2026-11-09: is_available 0인 방향은 정격(제한 없음), 둘 다 0이면 사용자 P 한도 끔.
			//   원래: 둘 다 0이면 아무것도 안 바꿈, 한쪽만 0이면 그 방향은 기존 값 유지 (처음 켤 때만 정격)]
			FOR u := 1 TO GVL_PARAM.UNIT_COUNT DO
				IF i_astUnitCfg[u].nPcs = p THEN
					_stUnit.astUnit[u].bPEnable	:= bCh OR bDis;
					IF bDis THEN
						_stUnit.astUnit[u].fPMax := fDis * MAX(i_astUnitCfg[u].fPRated, 0.0) / fSum;
					ELSE
						_stUnit.astUnit[u].fPMax := MAX(i_astUnitCfg[u].fPRated, 0.0);
					END_IF
					IF bCh THEN
						_stUnit.astUnit[u].fPMin := -(fCh * MAX(i_astUnitCfg[u].fPRated, 0.0) / fSum);
					ELSE
						_stUnit.astUnit[u].fPMin := -MAX(i_astUnitCfg[u].fPRated, 0.0);
					END_IF
				END_IF
			END_FOR
			bAny := TRUE;
		END_IF
	END_IF
END_FOR
IF bAny AND MEMCMP(ADR(_stUnit), ADR(iq_stUnitLimit), SIZEOF(_stUnit)) <> 0 THEN
	iq_stUnitLimit := _stUnit;
	M_Applied("EMS config: PCS 충·방전 전력 한도");
END_IF

(* BMS: SOC 최소·최대 → SOC 정책 (가장 엄격한 값). 값마다 숫자·0~100 먼저, 합친 설정은 F_SocLimitSetErr *)
_astBatBefore := _astBat;
_abBatRxBefore := _abBatRx;
bNewBat := FALSE;
FOR b := 1 TO GVL_PARAM.BMS_COUNT DO
	IF i_stCfg.anBatSeq[b] <> _anBatSeq[b] THEN
		_anBatSeq[b] := i_stCfg.anBatSeq[b];
		bBad := FALSE;
		// [UPS] SocMin·SocMax는 REAL (is_available 없음) → 둘 다 항상 검사
		bBad := NOT (F_RealOk(i_stCfg.astBat[b].SocMin) AND_THEN (i_stCfg.astBat[b].SocMin >= 0.0 AND i_stCfg.astBat[b].SocMin <= 100.0));
		IF NOT bBad THEN
			bBad := NOT (F_RealOk(i_stCfg.astBat[b].SocMax) AND_THEN (i_stCfg.astBat[b].SocMax >= 0.0 AND i_stCfg.astBat[b].SocMax <= 100.0));
		END_IF
		IF bBad THEN
			M_Reject(F_TxtNum("EMS config bat SOC 숫자·범위(0~100) 아님: BMS ", b));
		ELSE
			_astBat[b] := i_stCfg.astBat[b];
			_abBatRx[b] := TRUE;
			bNewBat := TRUE;
		END_IF
	END_IF
END_FOR
IF bNewBat THEN
	// [21번 수정 2026-11-09: is_available 0이면 기본값(하한 0 %, 상한 100 %)으로 보고 가장 엄격한 값을 고름. 기본값은 다른 BMS 값보다 엄격하지 않으므로
	//   값을 하나도 안 받은 BMS(빈 칸)는 결과에 영향이 없음. 원래: is_available 0은 계산에서 빼고, 하나도 없으면 기존 값 유지]
	fMin := SOC_MIN_DEFAULT;
	fMax := SOC_MAX_DEFAULT;
	FOR b := 1 TO GVL_PARAM.BMS_COUNT DO
		IF _abBatRx[b] AND_THEN _astBat[b].SocMin > fMin THEN		// [UPS] 받은 BMS만 (원래 SocMin.is_available <> 0 AND_THEN SocMin.value > fMin)
			fMin := _astBat[b].SocMin;
		END_IF
		IF _abBatRx[b] AND_THEN _astBat[b].SocMax < fMax THEN
			fMax := _astBat[b].SocMax;
		END_IF
	END_FOR
	_stSoc := iq_stSocLimit;
	_stSoc.fSocMin := fMin;
	_stSoc.fSocMax := fMax;
	_sErr := F_SocLimitSetErr(_stSoc);
	IF _sErr <> "" THEN
		_astBat := _astBatBefore;		// 이번에 받은 BMS 값은 버림 (다음 계산에 쓰지 않음)
		_abBatRx := _abBatRxBefore;
		M_Reject(WCONCAT("EMS config bat: ", _sErr));
	ELSIF MEMCMP(ADR(_stSoc), ADR(iq_stSocLimit), SIZEOF(_stSoc)) <> 0 THEN
		iq_stSocLimit := _stSoc;
		M_Applied("EMS config: SOC 상·하한");
	END_IF
END_IF

METHOD PRIVATE M_Reject
VAR_INPUT
	i_sText	: WSTRING(63);
END_VAR
q_bRejected	:= TRUE;
q_sRejected	:= i_sText;
q_nRejected	:= q_nRejected + 1;
END_METHOD

METHOD PRIVATE M_Applied
VAR_INPUT
	i_sText	: WSTRING(63);
END_VAR
q_bApplied	:= TRUE;
q_sApplied	:= i_sText;
q_nApplied	:= q_nApplied + 1;
END_METHOD

METHOD M_BuildEcho		// 실제 설정 → q_stEcho (MAIN이 설정 보호 뒤에 부름)
VAR_IN_OUT CONSTANT
	iq_stSocLimit	: ST_SocLimitSet;
	iq_stUnitLimit	: ST_UnitLimitSet;
END_VAR
VAR
	p			: UINT;
	u			: UINT;
	b			: UINT;
	bAll		: BOOL;
	bUnit		: BOOL;
	fMaxSum		: REAL;
	fMinSum		: REAL;
END_VAR
FOR p := 1 TO GVL_PARAM.PCS_COUNT DO
	bAll	:= TRUE;
	bUnit	:= FALSE;
	fMaxSum	:= 0.0;
	fMinSum	:= 0.0;
	FOR u := 1 TO GVL_PARAM.UNIT_COUNT DO
		IF i_astUnitCfg[u].nPcs = p THEN
			bUnit := TRUE;
			IF iq_stUnitLimit.astUnit[u].bPEnable AND F_RealOk(iq_stUnitLimit.astUnit[u].fPMax) AND F_RealOk(iq_stUnitLimit.astUnit[u].fPMin) THEN
				fMaxSum := fMaxSum + iq_stUnitLimit.astUnit[u].fPMax;
				fMinSum := fMinSum + iq_stUnitLimit.astUnit[u].fPMin;
			ELSE
				bAll := FALSE;
			END_IF
		END_IF
	END_FOR
	q_stEcho.astPcs[p - 1].DeviceId := UINT_TO_UDINT(p);	// 번호 1부터 [1부터 2026-11-10]
	IF bUnit AND bAll THEN
		q_stEcho.astPcs[p - 1].DisChargePowerLimit.value		:= DINT_TO_UDINT(MAX(F_RealToDint(fMaxSum), 0));
		q_stEcho.astPcs[p - 1].DisChargePowerLimit.is_available	:= 1;
		q_stEcho.astPcs[p - 1].ChargePowerLimit.value			:= DINT_TO_UDINT(MAX(F_RealToDint(-fMinSum), 0));
		q_stEcho.astPcs[p - 1].ChargePowerLimit.is_available		:= 1;
	ELSE
		q_stEcho.astPcs[p - 1].DisChargePowerLimit.value		:= 0;
		q_stEcho.astPcs[p - 1].DisChargePowerLimit.is_available	:= 0;
		q_stEcho.astPcs[p - 1].ChargePowerLimit.value			:= 0;
		q_stEcho.astPcs[p - 1].ChargePowerLimit.is_available		:= 0;
	END_IF
	q_stEcho.astPcs[p - 1].PvMarginRate.value			:= _stCfg.astPcs[p].PvMarginRate.value;	// 쓰지 않음: 받은 값, is_available 0
	q_stEcho.astPcs[p - 1].PvMarginRate.is_available	:= 0;
END_FOR
FOR b := 1 TO GVL_PARAM.BMS_COUNT DO
	q_stEcho.astBat[b - 1].DeviceId					:= UINT_TO_UDINT(b);	// 번호 1부터 [1부터 2026-11-10]
	q_stEcho.astBat[b - 1].SocMin					:= iq_stSocLimit.fSocMin;	// [UPS] REAL 형식 (원래 SocMin.value + is_available 1)
	q_stEcho.astBat[b - 1].SocMax					:= iq_stSocLimit.fSocMax;
END_FOR
END_METHOD

END_FUNCTION_BLOCK

// ---- 20_Module/Common/F_SocLimitSetErr.TcPOU
FUNCTION F_SocLimitSetErr : WSTRING(63)		// SOC 정책 설정 점검 ("" = 정상). FB_SocLimit.M_CheckSet과 FB_EmsConfigApply(EMS config 반영 전 검사)가 같이 씀 [9-21 수정 2026-11-04: FB_SocLimit.M_CheckSet에서 옮김]
VAR_INPUT
	i_stSet	: ST_SocLimitSet;
END_VAR

F_SocLimitSetErr := "";
IF NOT (F_RealOk(i_stSet.fSocMin) AND F_RealOk(i_stSet.fSocMax) AND F_RealOk(i_stSet.fBand) AND F_RealOk(i_stSet.fResumeMargin)) THEN	// [결함 13 수정 2026-11-04]
	F_SocLimitSetErr := "SOC 설정 숫자 아님";
ELSIF i_stSet.fSocMin < 0.0 OR i_stSet.fSocMax > 100.0 OR i_stSet.fSocMin >= i_stSet.fSocMax THEN
	F_SocLimitSetErr := "SOC 상·하한 (0 ≤ 하한 < 상한 ≤ 100)";
ELSIF i_stSet.fBand < 0.0 OR i_stSet.fSocMin + i_stSet.fBand > i_stSet.fSocMax - i_stSet.fBand THEN
	F_SocLimitSetErr := "감발 폭 fBand (0 이상, 상·하한 사이)";
ELSIF i_stSet.fResumeMargin < 0.0 OR i_stSet.fSocMin + i_stSet.fResumeMargin >= i_stSet.fSocMax - i_stSet.fResumeMargin THEN
	F_SocLimitSetErr := "재개 마진 fResumeMargin (0 이상, 상·하한 사이)";
END_IF

END_FUNCTION

// ---- 20_Module/Mqtt/FB_BrokerWatch.TcPOU
FUNCTION_BLOCK FB_BrokerWatch		// MQTT 브로커 끊김 감시 (PlcTask, MAIN이 부름) [9번 수정 2026-11-09: 추가 — 14번 탭 9번 결정]
// - 감시: i_stSet.eBroker로 고른 브로커가 쓰는 브로커(MQTT_SET bUse)일 때만. 접속 상태는 PRG_Mqtt가 GVL_IF.g_abBrokerConn에 올림 (구독 클라이언트 기준)
// - 끊김: 접속이 i_stSet.tLostDelay 넘게 이어서 끊기면 q_bLost (알람 '브로커 끊김', 접속하면 해소). PMS 시작 직후 접속 전도 끊김으로 셈
// - Manual 전환: 끊김 동안 한 번만 q_bToManual (1스캔) → MAIN이 운전 모드 요청(g_aeOpMode)을 모두 Manual로. 끊긴 동안 운전원이 Auto로 되돌려도 다시 바꾸지 않음.
//   다시 접속하면(q_bLost 해소) 다시 무장 → 다음 끊김에 다시 한 번
// - 이중화: Active PLC만 전환 요청 (대기 PLC의 운전 모드 요청은 Active 값으로 동기화됨). 끊긴 동안 Active가 되면 그때 한 번
VAR_INPUT
	i_stSet			: ST_BrokerWatchSet;
	i_abUse			: ARRAY[1..3] OF BOOL;	// 쓰는 브로커 (GVL_IF.g_abBrokerUse, 1 Cloud, 2 Local, 3 Azure)
	i_abConnected	: ARRAY[1..3] OF BOOL;	// 접속됨 (GVL_IF.g_abBrokerConn)
	i_bActive		: BOOL;					// 이 PLC가 Active (GVL_IF.g_bRedActive. 이중화를 안 쓰면 항상 TRUE)
END_VAR
VAR_OUTPUT
	q_bWatch		: BOOL;			// 감시 중 (고른 브로커를 씀)
	q_bLost			: BOOL;			// 끊김 확정 (알람)
	q_bToManual		: BOOL;			// 이번 스캔에 Manual 전환 요청 (1스캔)
	q_sBroker		: WSTRING(15);	// 고른 브로커 이름 (로그)
	q_sDelay		: WSTRING(31);	// 판정 시간 글자 (로그)
END_VAR
VAR
	_tonLost		: TON;
	_bDone			: BOOL;			// 이번 끊김에서 전환 요청을 냄 (접속하면 지움)
	_n				: INT;			// 고른 브로커 칸 (0 = 범위 밖)
END_VAR

CASE i_stSet.eBroker OF
	E_MqttBroker.Cloud:	_n := 1;	q_sBroker := "Cloud";
	E_MqttBroker.Local:	_n := 2;	q_sBroker := "Local";
	E_MqttBroker.Azure:	_n := 3;	q_sBroker := "Azure";
ELSE
	_n := 0;	q_sBroker := "?";
END_CASE
q_sDelay := WCONCAT(TO_WSTRING(TIME_TO_UDINT(i_stSet.tLostDelay) / 1000), " s");

q_bWatch := FALSE;
IF _n >= 1 AND _n <= 3 THEN
	q_bWatch := i_abUse[_n];
END_IF
IF q_bWatch THEN
	_tonLost(IN := NOT i_abConnected[_n], PT := i_stSet.tLostDelay);
ELSE
	_tonLost(IN := FALSE);
END_IF
q_bLost := _tonLost.Q;

q_bToManual := q_bLost AND NOT _bDone AND i_bActive;
IF q_bToManual THEN
	_bDone := TRUE;
END_IF
IF NOT q_bLost THEN
	_bDone := FALSE;		// 다시 접속: 다음 끊김에 다시 한 번
END_IF

END_FUNCTION_BLOCK

// ---- 20_Module/Virtual/PRG_SimLink.TcPOU
PROGRAM PRG_SimLink		// 가상 장비끼리 연결 (사무실 시험 전용)
VAR_TEMP
	u			: UINT;
	p			: UINT;
	stUnit		: ST_UnitState;
	fP			: REAL;
	fQ			: REAL;
	b			: UINT;
	afPBat		: ARRAY[1..GVL_PARAM.BAT_COUNT] OF REAL;	// kW, 배터리 그룹(DC 버스)마다 유닛 P 합
END_VAR

(* 실제 현장에서 전기가 이어 주는 것을 흉내 냄: PCS 출력 → 배터리 SOC, 접속점 계측
   - 가상 PCS 여러 대(GVL_SITE.g_aipPcs) → 배터리 그룹마다 그 그룹 BMS (GVL_SITE.BMS_CFG), 계측기1 하나 기준
   - BMS를 늘리거나 줄이면 아래 BMS 줄도 같이 맞춤
   - 현장 빌드: GVL_SITE의 장비를 실제 드라이버로 바꾸고, MAIN의 PRG_SimLink() 호출과 Virtual 폴더 삭제 *)
fP := 0;
fQ := 0;
FOR b := 1 TO GVL_PARAM.BAT_COUNT DO
	afPBat[b] := 0;
END_FOR
FOR u := 1 TO GVL_PARAM.UNIT_COUNT DO
	p := GVL_SITE.UNIT_CFG[u].nPcs;
	IF p >= 1 AND p <= GVL_PARAM.PCS_COUNT THEN
		IF GVL_SITE.g_aipPcs[p] <> 0 THEN
			stUnit	:= GVL_SITE.g_aipPcs[p].M_GetUnitState(GVL_SITE.UNIT_CFG[u].nSub);
			fP		:= fP + stUnit.stP.fValue;
			fQ		:= fQ + stUnit.stQ.fValue;
			b		:= GVL_SITE.UNIT_CFG[u].nBatGroup;
			IF b >= 1 AND b <= GVL_PARAM.BAT_COUNT THEN
				afPBat[b] := afPBat[b] + stUnit.stP.fValue;
			END_IF
		END_IF
	END_IF
END_FOR
// BMS1: physical-map driver has no simulated power input.
// BMS2: physical-map driver has no simulated power input.
// BMS3: physical-map driver has no simulated power input.
GVL_SITE.g_fbMeter1.i_fP	:= fP;
GVL_SITE.g_fbMeter1.i_fQ	:= fQ;

END_PROGRAM

// ---- 99_Test/PRG_TestCtrlMode.TcPOU
PROGRAM PRG_TestCtrlMode		// 제어 모드 자동 시험 (GVL_SITE.TEST_MODE일 때 MAIN이 부름). 실제 제어와 따로 둔 인스턴스만 씀 (장비 지령에 영향 없음)
// 온라인에서 bDone = TRUE가 되면 fbTally.q_nPass·q_nFail, 실패하면 fbTally.q_anFail(실패한 시험 번호)을 봄. bRestart := TRUE로 다시 돌림
// 1~16: 스케줄 모드 단위 시험 (한 스캔). 20~32: 관리자 전환 시험 (여러 스캔, 약 3 s)
VAR
	bRestart	: BOOL;			// TRUE로 쓰면 처음부터 다시
	bDone		: BOOL;			// 시험 끝
	nStep		: UINT;
	fbTally		: FB_TestTally;
	fbSched		: FB_CmSchedule		:= (i_nModuleId := 9001, i_sName := 'TestSched');
	fbConst		: FB_CmConstPower	:= (i_nModuleId := 9002, i_sName := 'TestConst');
	fbMgr		: FB_CtrlModeMgr	:= (i_nModuleId := 9000, i_sName := 'TestMgr');
	aipMode		: ARRAY[1..GVL_PARAM.CTRL_MODE_COUNT] OF I_ControlMode;	// 1 = 정출력 50 kW, 2 = 스케줄
	stCommon	: ST_CmCommonSet;
	stTable		: ST_CmScheduleSet;
	stView		: ST_CtrlModeView;
	stOut		: ST_CtrlModeOut;
	stMgrOut	: ST_SourceOutput;
	stReg		: ST_SourceReg := (bEnable := TRUE, nGrade := 1, ePowerMode := E_SourceMode.Auto, nGroup := 0, tExpire := T#10S);
	tonWait		: TON;
	wsTmp		: WSTRING(63);
END_VAR

IF bRestart THEN
	bRestart	:= FALSE;
	bDone		:= FALSE;
	nStep		:= 0;
END_IF

CASE nStep OF
	0:	// 준비 + 스케줄 단위 시험 (한 스캔)
		fbTally.M_Reset();
		A_Setup();
		A_UnitSchedule();
		fbMgr.i_nModeReq := 2;
		nStep := 10;

	10:	// 관리자: 모드 없음 → 스케줄(2). 켜진 모드가 없으므로 바로 진입
		A_CycleMgr();
		fbTally.M_Check(i_nId := 20, i_bOk := fbMgr.q_nActive = 2 AND fbMgr.q_eStep = E_CtrlModeStep.Active);
		fbTally.M_Check(i_nId := 21, i_bOk := stMgrOut.bPSetActive AND ABS(stMgrOut.fPSet - 200.0) < 0.01);
		fbMgr.i_nModeReq := 1;
		nStep := 11;

	11:	// 정출력(1) 요청 첫 스캔: 이전 모드 끝, 출력 0으로 전환 중
		A_CycleMgr();
		fbTally.M_Check(i_nId := 22, i_bOk := fbMgr.q_eStep = E_CtrlModeStep.Leaving AND fbMgr.q_nActive = 0 AND fbMgr.q_nTarget = 1);
		fbTally.M_Check(i_nId := 23, i_bOk := stMgrOut.bPSetActive AND ABS(stMgrOut.fPSet) < 0.01);
		nStep := 12;

	12:	// tZeroDelay(1 s) 뒤 정출력 진입
		A_CycleMgr();
		tonWait(IN := TRUE, PT := T#3S);
		IF fbMgr.q_eStep = E_CtrlModeStep.Active OR tonWait.Q THEN
			fbTally.M_Check(i_nId := 24, i_bOk := fbMgr.q_nActive = 1 AND ABS(stMgrOut.fPSet - 50.0) < 0.01);
			fbTally.M_Check(i_nId := 25, i_bOk := tonWait.ET >= T#900MS AND NOT tonWait.Q);
			tonWait(IN := FALSE);
			fbMgr.i_nModeReq := 9;
			nStep := 13;
		END_IF

	13:	// 없는 칸(9) → BadSlot, 지금 모드 유지
		A_CycleMgr();
		fbTally.M_Check(i_nId := 26, i_bOk := fbMgr.q_eRefuse = E_CtrlModeRefuse.BadSlot AND fbMgr.q_nActive = 1);
		stView.stTime.bValid	:= FALSE;
		fbMgr.i_nModeReq		:= 2;
		nStep := 14;

	14:	// 시각 무효 → 스케줄 진입 거부 (NotReady, 이유 NO_TIME), 정출력 유지
		A_CycleMgr();
		fbTally.M_Check(i_nId := 27, i_bOk := fbMgr.q_eRefuse = E_CtrlModeRefuse.NotReady AND fbMgr.q_nRefuseReason = GVL_CM_RSN.NO_TIME AND fbMgr.q_nActive = 1);
		fbTally.M_Check(i_nId := 28, i_bOk := ABS(stMgrOut.fPSet - 50.0) < 0.01);
		stView.stTime.bValid	:= TRUE;
		fbMgr.i_bRetry			:= TRUE;		// 같은 요청(2)을 다시
		nStep := 15;

	15:	// 재시도 → 전환 시작
		A_CycleMgr();
		fbTally.M_Check(i_nId := 29, i_bOk := fbMgr.q_eStep = E_CtrlModeStep.Leaving AND fbMgr.q_nTarget = 2 AND NOT fbMgr.i_bRetry);
		nStep := 16;

	16:	// 스케줄 진입
		A_CycleMgr();
		tonWait(IN := TRUE, PT := T#3S);
		IF fbMgr.q_eStep = E_CtrlModeStep.Active OR tonWait.Q THEN
			fbTally.M_Check(i_nId := 30, i_bOk := fbMgr.q_nActive = 2 AND ABS(stMgrOut.fPSet - 200.0) < 0.01);
			tonWait(IN := FALSE);
			fbMgr.i_nModeReq := 0;
			nStep := 17;
		END_IF

	17:	// 모드 없음(0) → 출력 0 뒤 지령 없음
		A_CycleMgr();
		tonWait(IN := TRUE, PT := T#3S);
		IF fbMgr.q_eStep = E_CtrlModeStep.Idle OR tonWait.Q THEN
			fbTally.M_Check(i_nId := 31, i_bOk := fbMgr.q_eStep = E_CtrlModeStep.Idle AND fbMgr.q_nActive = 0 AND NOT stMgrOut.bPSetActive);
			tonWait(IN := FALSE);
			// 설정 점검: 시작 > 끝인 칸이 있으면 관리자가 모드의 오류 문구를 올림
			stTable.astSlot[2, 3, 5].nStart	:= 1500;
			stTable.astSlot[2, 3, 5].nEnd	:= 1400;
			fbSched.i_stTable := stTable;
			wsTmp := fbMgr.M_CheckSet();
			fbTally.M_Check(i_nId := 32, i_bOk := wsTmp <> "");
			stTable.astSlot[2, 3, 5].nStart	:= 0;
			stTable.astSlot[2, 3, 5].nEnd	:= 0;
			fbSched.i_stTable := stTable;
			wsTmp := fbMgr.M_CheckSet();
			fbTally.M_Check(i_nId := 33, i_bOk := wsTmp = "");
			nStep := 99;
		END_IF

	99:
		bDone := TRUE;
END_CASE

ACTION A_Setup:
// 모드 등록·설정
aipMode[1]	:= fbConst;
aipMode[2]	:= fbSched;
fbConst.i_stSet.fPSet	:= 50.0;
fbConst.i_stSet.bQSet	:= FALSE;
fbConst.i_stSet.tDuration	:= T#0S;
// 공통 설정: 기본값(방전 08:00~22:00, 일요일 금지, 역송 여유 10 kW·0.95) + 7월 14일 휴일
stCommon.abHoliday[7, 14]	:= TRUE;
// 시간표: 여름(0) 월요일(1), 일요일(0)
stTable.astSlot[0, 1, 1].nStart := 100;		stTable.astSlot[0, 1, 1].nEnd := 600;		stTable.astSlot[0, 1, 1].fP := -300.0;	// 충전
stTable.astSlot[0, 1, 2].nStart := 1000;	stTable.astSlot[0, 1, 2].nEnd := 1200;		stTable.astSlot[0, 1, 2].fP := 200.0;	// 방전
stTable.astSlot[0, 1, 3].nStart := 1100;	stTable.astSlot[0, 1, 3].nEnd := 1130;		stTable.astSlot[0, 1, 3].fP := 400.0;	// 겹침: 번호 큰 칸
stTable.astSlot[0, 1, 4].nStart := 2300;	stTable.astSlot[0, 1, 4].nEnd := 2400;		stTable.astSlot[0, 1, 4].fP := 100.0;	// 방전 허용 시간 밖
stTable.astSlot[0, 0, 1].nStart := 1000;	stTable.astSlot[0, 0, 1].nEnd := 1200;		stTable.astSlot[0, 0, 1].fP := 200.0;	// 일요일
fbSched.i_stCommon	:= stCommon;
fbSched.i_stTable	:= stTable;
// 관리자: 기본 설정 (전환 때 1 s 출력 0, 대체 모드 없음)
fbMgr.i_stSet.bZeroOnSwitch	:= TRUE;
fbMgr.i_stSet.tZeroDelay	:= T#1S;
fbMgr.i_stSet.nFallback		:= 0;
fbMgr.i_bRetry				:= FALSE;
A_ViewBase();
END_ACTION

ACTION A_ViewBase:
// 기준 상황: 2026-07-13 월요일 10:30:00, 가용 유닛 1, 가용 출력 1000 kW, 수전 1000 kW (접속점 P = -1000), ESS 출력 0
stView.stTime.bValid		:= TRUE;
stView.stTime.nYear			:= 2026;
stView.stTime.nMonth		:= 7;
stView.stTime.nDay			:= 13;
stView.stTime.nDayOfWeek	:= 1;
stView.stTime.nHour			:= 10;
stView.stTime.nMinute		:= 30;
stView.stTime.nSecond		:= 0;
stView.stGroup.nUnitAvail	:= 1;
stView.stGroup.fPRatedAvail	:= 1000.0;
stView.stGroup.fPOut		:= 0.0;
stView.stGroup.stPcc.stMeas.stP.bValid	:= TRUE;
stView.stGroup.stPcc.stMeas.stP.fValue	:= -1000.0;
END_ACTION

ACTION A_UnitSchedule:
fbSched.M_Enter(i_stView := stView);

// 1) 03:00 충전 칸 → -300
A_ViewBase();
stView.stTime.nHour := 3;	stView.stTime.nMinute := 0;
stOut := fbSched.M_Calc(i_stView := stView);
fbTally.M_Check(i_nId := 1, i_bOk := ABS(stOut.fPSet + 300.0) < 0.01 AND fbSched.q_nSlot = 1 AND fbSched.q_nState = 0);

// 2) 10:30 방전 칸 → 200
A_ViewBase();
stOut := fbSched.M_Calc(i_stView := stView);
fbTally.M_Check(i_nId := 2, i_bOk := ABS(stOut.fPSet - 200.0) < 0.01 AND fbSched.q_nSlot = 2 AND fbSched.q_nState = 0);

// 3) 11:15 겹친 칸 → 번호 큰 칸 400
A_ViewBase();
stView.stTime.nHour := 11;	stView.stTime.nMinute := 15;
stOut := fbSched.M_Calc(i_stView := stView);
fbTally.M_Check(i_nId := 3, i_bOk := ABS(stOut.fPSet - 400.0) < 0.01 AND fbSched.q_nSlot = 3);

// 4) 12:00 = 끝 시각 (미포함) → 칸 없음 0, 지령은 냄
A_ViewBase();
stView.stTime.nHour := 12;	stView.stTime.nMinute := 0;
stOut := fbSched.M_Calc(i_stView := stView);
fbTally.M_Check(i_nId := 4, i_bOk := stOut.bPSetActive AND ABS(stOut.fPSet) < 0.01 AND fbSched.q_nSlot = 0 AND fbSched.q_nState = GVL_CM_RSN.NO_SLOT);

// 5) 23:30 방전 칸이지만 방전 허용 시간 밖 → 0
A_ViewBase();
stView.stTime.nHour := 23;
stOut := fbSched.M_Calc(i_stView := stView);
fbTally.M_Check(i_nId := 5, i_bOk := ABS(stOut.fPSet) < 0.01 AND fbSched.q_nSlot = 4 AND fbSched.q_nState = GVL_CM_RSN.DIS_TIME);

// 6) 일요일 10:30 방전 칸 → 일요일 방전 금지로 0
A_ViewBase();
stView.stTime.nDayOfWeek := 0;	stView.stTime.nDay := 12;
stOut := fbSched.M_Calc(i_stView := stView);
fbTally.M_Check(i_nId := 6, i_bOk := ABS(stOut.fPSet) < 0.01 AND fbSched.q_nSlot = 1 AND fbSched.q_nState = GVL_CM_RSN.DIS_TIME);

// 7) 역송 방지: 수전 150 kW → 부하 150, 가능 140 → 140 × 0.95 = 133
A_ViewBase();
stView.stGroup.stPcc.stMeas.stP.fValue := -150.0;
stOut := fbSched.M_Calc(i_stView := stView);
fbTally.M_Check(i_nId := 7, i_bOk := ABS(stOut.fPSet - 133.0) < 0.01 AND fbSched.q_nState = GVL_CM_RSN.REV_LIMIT);

// 8) 접속점 계측 무효 → 방전 0
A_ViewBase();
stView.stGroup.stPcc.stMeas.stP.bValid := FALSE;
stOut := fbSched.M_Calc(i_stView := stView);
fbTally.M_Check(i_nId := 8, i_bOk := ABS(stOut.fPSet) < 0.01 AND fbSched.q_nState = GVL_CM_RSN.NO_PCC);

// 9) 휴일 (7월 14일) → 0
A_ViewBase();
stView.stTime.nDay := 14;	stView.stTime.nDayOfWeek := 2;
stOut := fbSched.M_Calc(i_stView := stView);
fbTally.M_Check(i_nId := 9, i_bOk := ABS(stOut.fPSet) < 0.01 AND fbSched.q_nState = GVL_CM_RSN.HOLIDAY);

// 10) 시각 무효 → 0, 진입 거부 이유 NO_TIME
A_ViewBase();
stView.stTime.bValid := FALSE;
stOut := fbSched.M_Calc(i_stView := stView);
fbTally.M_Check(i_nId := 10, i_bOk := ABS(stOut.fPSet) < 0.01 AND fbSched.q_nState = GVL_CM_RSN.NO_TIME AND fbSched.M_CheckEnter(i_stView := stView) = GVL_CM_RSN.NO_TIME);

// 11) 1월 = 겨울(2): 겨울 시간표가 비어 칸 없음
A_ViewBase();
stView.stTime.nMonth := 1;
stOut := fbSched.M_Calc(i_stView := stView);
fbTally.M_Check(i_nId := 11, i_bOk := fbSched.q_nSeason = 2 AND fbSched.q_nState = GVL_CM_RSN.NO_SLOT);

// 12) ESS 충전 중 역송 방지: 수전 500, ESS -300 → 부하 200, 가능 190 → 180.5
A_ViewBase();
stView.stGroup.stPcc.stMeas.stP.fValue := -500.0;
stView.stGroup.fPOut := -300.0;
stOut := fbSched.M_Calc(i_stView := stView);
fbTally.M_Check(i_nId := 12, i_bOk := ABS(stOut.fPSet - 180.5) < 0.01 AND fbSched.q_nState = GVL_CM_RSN.REV_LIMIT);

// 13) 진입 검사: 정상이면 0
A_ViewBase();
fbTally.M_Check(i_nId := 13, i_bOk := fbSched.M_CheckEnter(i_stView := stView) = 0);

// 14) 설정 점검: 시작 > 끝인 칸 → 오류 문구, 되돌리면 정상
stTable.astSlot[1, 4, 2].nStart := 1300;	stTable.astSlot[1, 4, 2].nEnd := 1200;
fbSched.i_stTable := stTable;
wsTmp := fbSched.M_CheckSet();
fbTally.M_Check(i_nId := 14, i_bOk := wsTmp <> "");
stTable.astSlot[1, 4, 2].nStart := 0;		stTable.astSlot[1, 4, 2].nEnd := 0;
fbSched.i_stTable := stTable;
wsTmp := fbSched.M_CheckSet();
fbTally.M_Check(i_nId := 15, i_bOk := wsTmp = "");

// 16) 방전 허용 시간을 끄면 23:30 방전 칸 100
stCommon.stDis.bUse := FALSE;
fbSched.i_stCommon := stCommon;
A_ViewBase();
stView.stTime.nHour := 23;
stOut := fbSched.M_Calc(i_stView := stView);
fbTally.M_Check(i_nId := 16, i_bOk := ABS(stOut.fPSet - 100.0) < 0.01 AND fbSched.q_nState = 0);
stCommon.stDis.bUse := TRUE;
fbSched.i_stCommon := stCommon;

// 17) 진입 검사: 가용 유닛 없음 → NO_UNIT
A_ViewBase();
stView.stGroup.nUnitAvail := 0;
fbTally.M_Check(i_nId := 17, i_bOk := fbSched.M_CheckEnter(i_stView := stView) = GVL_CM_RSN.NO_UNIT);

fbSched.M_Exit();
A_ViewBase();
END_ACTION

ACTION A_CycleMgr:
// 관리자 한 스캔 (FB_SourceHub가 하는 것처럼 M_Cycle을 부름)
fbMgr.i_aipMode	:= aipMode;
fbMgr.i_stTime	:= stView.stTime;
fbMgr.M_Cycle(i_stReg := stReg, i_stView := stView.stGroup);
stMgrOut := fbMgr.Output;
END_ACTION

END_PROGRAM

// ---- 99_Test/FB_TestTally.TcPOU
FUNCTION_BLOCK FB_TestTally		// 시험 결과 세기: 통과·실패 수와 실패한 시험 번호
VAR_OUTPUT
	q_nPass		: UINT;
	q_nFail		: UINT;
	q_anFail	: ARRAY[1..32] OF UINT;		// 실패한 시험 번호 (앞에서부터)
END_VAR

METHOD M_Reset
VAR
	nI	: UINT;
END_VAR
q_nPass := 0;
q_nFail := 0;
FOR nI := 1 TO 32 DO
	q_anFail[nI] := 0;
END_FOR
END_METHOD

METHOD M_Check : BOOL
VAR_INPUT
	i_nId	: UINT;		// 시험 번호
	i_bOk	: BOOL;
END_VAR
IF i_bOk THEN
	q_nPass := q_nPass + 1;
ELSE
	q_nFail := q_nFail + 1;
	IF q_nFail <= 32 THEN
		q_anFail[q_nFail] := i_nId;
	END_IF
END_IF
M_Check := i_bOk;
END_METHOD

END_FUNCTION_BLOCK

// ---- 20_Module/ControlMode/FB_CmSchedule.TcPOU
FUNCTION_BLOCK FB_CmSchedule EXTENDS FB_CmTariffBase		// 제어 모드: 스케줄 (Messis SCHEDULE_MODE). 계절·요일 시간표의 P를 냄
// 맞는 칸 없음·휴일·시각 무효 → 0. 충전(-)은 그대로, 방전(+)은 방전 허용 시간·역송 방지 (공통 설정). 칸은 자정을 넘지 않음
VAR_INPUT
	i_stTable	: ST_CmScheduleSet;		// 시간표 (A_PassModuleSet이 GVL_PERSIST.g_stModuleSet.stCmSchedule을 매 스캔 넘김)
END_VAR

METHOD M_Calc : ST_CtrlModeOut
VAR_INPUT
	i_stView	: ST_CtrlModeView;
END_VAR
VAR
	fP		: REAL;
	nRsn	: UINT;
END_VAR
fP := 0.0;
IF M_Begin(i_stView := i_stView) THEN
	M_SchedLookup(i_stTime := i_stView.stTime, iq_stTable := i_stTable);
	fP			:= M_SchedOut(i_stView := i_stView, q_nRsn => nRsn);
	q_nState	:= nRsn;
END_IF
M_Calc := M_Finish(i_fP := fP);
END_METHOD

METHOD M_CheckSet : WSTRING(63)
M_CheckSet := SUPER^.M_CheckSet();
IF M_CheckSet = "" THEN
	M_CheckSet := M_CheckTable(iq_stTable := i_stTable);
END_IF
END_METHOD

END_FUNCTION_BLOCK

// ---- 20_Module/ControlMode/FB_CmTariffBase.TcPOU
FUNCTION_BLOCK ABSTRACT FB_CmTariffBase EXTENDS FB_CtrlModeBase		// 요금제 기반 제어 모드 공통 바탕 (스케줄·피크컷·통합). 같은 계산은 여기 메서드 하나만 씀
// 휴일·계절·방전 허용 시간·역송 방지·시간표 조회·잔량 방전·자동 충전. 상태·이유 코드는 GVL_CM_RSN
// 파생 FB: M_Calc에서 M_Begin으로 시작 → 계산 → M_Finish로 끝냄
VAR_INPUT
	i_stCommon	: ST_CmCommonSet;	// 공통 설정 (A_PassModuleSet이 GVL_PERSIST.g_stModuleSet.stCmCommon을 매 스캔 넘김)
END_VAR
VAR_OUTPUT
	q_nState	: UINT;		// 0 = 정상, 그 외 = GVL_CM_RSN (M_ReasonText)
	q_fOutP		: REAL;		// 이번 스캔에 낸 P (kW, 방전 +)
	q_nSeason	: UINT;		// 지금 계절 (0 여름, 1 봄·가을, 2 겨울)
	q_nSlot		: UINT;		// 맞는 시간표 칸 (0 = 없음, 시간표를 쓰는 모드만)
	q_fSlotP	: REAL;		// 그 칸 값 (kW)
END_VAR

METHOD M_CheckEnter : UINT
VAR_INPUT
	i_stView	: ST_CtrlModeView;
END_VAR
M_CheckEnter := 0;
IF NOT M_TimeOk(i_stTime := i_stView.stTime) THEN
	M_CheckEnter := GVL_CM_RSN.NO_TIME;
ELSIF i_stView.stGroup.nUnitAvail = 0 THEN
	M_CheckEnter := GVL_CM_RSN.NO_UNIT;
END_IF
END_METHOD

METHOD PROTECTED M_Begin : BOOL		// 스캔 시작: 출력 칸을 비우고 계절을 셈. 시각이 맞고 휴일이 아니면 TRUE (FALSE면 q_nState에 이유, 0을 냄)
VAR_INPUT
	i_stView	: ST_CtrlModeView;
END_VAR
q_nState	:= 0;
q_fOutP		:= 0.0;
q_nSlot		:= 0;
q_fSlotP	:= 0.0;
M_Begin		:= FALSE;
IF NOT M_TimeOk(i_stTime := i_stView.stTime) THEN
	q_nState := GVL_CM_RSN.NO_TIME;
ELSE
	q_nSeason := i_stCommon.anSeasonOfMonth[i_stView.stTime.nMonth];
	IF q_nSeason > 2 THEN
		q_nSeason := 0;		// M_CheckSet이 막지만 배열 범위 보호
	END_IF
	IF i_stCommon.abHoliday[i_stView.stTime.nMonth, i_stView.stTime.nDay] THEN
		q_nState := GVL_CM_RSN.HOLIDAY;
	ELSE
		M_Begin := TRUE;
	END_IF
END_IF
END_METHOD

METHOD PROTECTED M_Finish : ST_CtrlModeOut		// 스캔 끝: P를 지령으로 냄 (0이어도 냄: 등급이 낮은 지령원으로 넘어가지 않게). Q는 내지 않음
VAR_INPUT
	i_fP		: REAL;		// kW, 방전 +
END_VAR
q_fOutP					:= i_fP;
M_Finish.bPSetActive	:= TRUE;
M_Finish.fPSet			:= i_fP;
M_Finish.bQSetActive	:= FALSE;
M_Finish.fQSet			:= 0.0;
M_Finish.bExitReq		:= FALSE;
M_Finish.nReason		:= 0;
END_METHOD

METHOD PROTECTED M_TimeOk : BOOL		// 시각이 유효하고 배열 번호로 쓸 수 있는 범위
VAR_INPUT
	i_stTime	: ST_LocalTime;
END_VAR
M_TimeOk := i_stTime.bValid AND i_stTime.nMonth >= 1 AND i_stTime.nMonth <= 12
	AND i_stTime.nDay >= 1 AND i_stTime.nDay <= 31 AND i_stTime.nDayOfWeek <= 6;
END_METHOD

METHOD PROTECTED M_DisAllowed : BOOL		// 지금 방전해도 되는 시간인가 (공통 설정 stDis)
VAR_INPUT
	i_stTime	: ST_LocalTime;
END_VAR
M_DisAllowed := TRUE;
IF i_stCommon.stDis.bUse THEN
	M_DisAllowed := F_InHhmmWindow(i_nNow := F_TimeHhmm(i_stTime := i_stTime), i_nStart := i_stCommon.stDis.nStart, i_nEnd := i_stCommon.stDis.nEnd)
		AND (i_stTime.nDayOfWeek <> 0 OR i_stCommon.stDis.bSunday);
END_IF
END_METHOD

METHOD PROTECTED M_NoReverse : REAL		// 역송 방지: 방전 요청을 (부하 − 여유) 안으로 줄임 (공통 설정 stNoRev). 충전·0은 그대로
VAR_INPUT
	i_fReq		: REAL;		// kW, 방전 +
	i_stView	: ST_CtrlModeView;
END_VAR
VAR_OUTPUT
	q_nRsn		: UINT;		// 0 = 그대로, GVL_CM_RSN.REV_LIMIT = 줄임, GVL_CM_RSN.NO_PCC = 계측 무효로 0
END_VAR
VAR
	fLoad		: REAL;		// 부하 = ESS가 없을 때의 수전
	fAvail		: REAL;		// 역송 없이 방전할 수 있는 양
END_VAR
M_NoReverse	:= i_fReq;
q_nRsn		:= 0;
IF i_fReq > 0.0 AND i_stCommon.stNoRev.bUse THEN
	IF i_stView.stGroup.stPcc.stMeas.stP.bValid THEN
		// 접속점 P는 공급(역송) +, 수전 -. 부하 = ESS 출력 − 접속점 공급 (충전 중·역송 중에도 맞음)
		fLoad	:= MAX(i_stView.stGroup.fPOut - i_stView.stGroup.stPcc.stMeas.stP.fValue, 0.0);
		fAvail	:= MAX(fLoad - i_stCommon.stNoRev.fMargin, 0.0);
		IF i_fReq > fAvail THEN
			M_NoReverse	:= fAvail * i_stCommon.stNoRev.fScale;
			q_nRsn		:= GVL_CM_RSN.REV_LIMIT;
		END_IF
	ELSE
		M_NoReverse	:= 0.0;
		q_nRsn		:= GVL_CM_RSN.NO_PCC;
	END_IF
END_IF
END_METHOD

METHOD PROTECTED M_SchedLookup : BOOL		// 시간표에서 지금 맞는 칸 (번호가 큰 칸 우선). 찾으면 TRUE, q_nSlot·q_fSlotP에 씀. M_Begin 뒤에 부름 (계절)
VAR_INPUT
	i_stTime	: ST_LocalTime;
END_VAR
VAR_IN_OUT CONSTANT
	iq_stTable	: ST_CmScheduleSet;
END_VAR
VAR
	nNow		: UINT;
	k			: UINT;
END_VAR
nNow		:= F_TimeHhmm(i_stTime := i_stTime);
q_nSlot		:= 0;
q_fSlotP	:= 0.0;
FOR k := 1 TO GVL_PARAM.SCHED_SLOT_COUNT DO
	IF F_InHhmmWindow(i_nNow := nNow, i_nStart := iq_stTable.astSlot[q_nSeason, i_stTime.nDayOfWeek, k].nStart, i_nEnd := iq_stTable.astSlot[q_nSeason, i_stTime.nDayOfWeek, k].nEnd) THEN
		q_nSlot		:= k;
		q_fSlotP	:= iq_stTable.astSlot[q_nSeason, i_stTime.nDayOfWeek, k].fP;
	END_IF
END_FOR
M_SchedLookup := q_nSlot <> 0;
END_METHOD

METHOD PROTECTED M_SchedOut : REAL		// 시간표 값 → 낼 값: 칸 없음 0, 충전 그대로, 방전은 방전 허용 시간·역송 방지 (스케줄·통합 모드 공통)
VAR_INPUT
	i_stView	: ST_CtrlModeView;
END_VAR
VAR_OUTPUT
	q_nRsn		: UINT;		// 0 = 칸 값 그대로, 그 외 GVL_CM_RSN
END_VAR
q_nRsn		:= 0;
M_SchedOut	:= 0.0;
IF q_nSlot = 0 THEN
	q_nRsn := GVL_CM_RSN.NO_SLOT;
ELSIF q_fSlotP > 0.0 THEN
	IF M_DisAllowed(i_stTime := i_stView.stTime) THEN
		M_SchedOut := M_NoReverse(i_fReq := q_fSlotP, i_stView := i_stView, q_nRsn => q_nRsn);
	ELSE
		q_nRsn := GVL_CM_RSN.DIS_TIME;
	END_IF
ELSE
	M_SchedOut := q_fSlotP;		// 충전 (또는 0)
END_IF
END_METHOD

METHOD PROTECTED M_RemainDis : REAL		// 잔량 방전량 (kW): (지금 에너지 − 하한 SOC 에너지)를 끝 시각까지 고르게. 가용 출력 상한. 역송 방지 전
VAR_INPUT
	i_stView	: ST_CtrlModeView;
	i_stWin		: ST_CmWindowSet;	// nEnd, fSoc = 남길 하한
END_VAR
VAR_OUTPUT
	q_bNoCap	: BOOL;		// 용량·SOC 무효
END_VAR
VAR
	nMin		: UINT;
	fE			: REAL;		// kWh
END_VAR
M_RemainDis	:= 0.0;
q_bNoCap	:= i_stView.stGroup.fCapacity <= 0.0 OR NOT i_stView.stGroup.stSocAvg.bValid;
IF NOT q_bNoCap THEN
	nMin	:= F_MinutesTo(i_nNow := F_TimeHhmm(i_stTime := i_stView.stTime), i_nEnd := i_stWin.nEnd);
	fE		:= i_stView.stGroup.fCapacity * (i_stView.stGroup.stSocAvg.fValue - i_stWin.fSoc) / 100.0;
	IF nMin > 0 AND fE > 0.0 THEN
		M_RemainDis := MIN(fE * 60.0 / UINT_TO_REAL(nMin), i_stView.stGroup.fPRatedAvail);
	END_IF
END_IF
END_METHOD

METHOD PROTECTED M_AutoChg : REAL		// 자동 충전량 (kW, 양수): (목표 SOC 에너지 − 지금 에너지)를 끝 시각까지 + 1 kW, 최소 10 kW, 가용 출력 상한
VAR_INPUT
	i_stView	: ST_CtrlModeView;
	i_stWin		: ST_CmWindowSet;	// nEnd, fSoc = 채울 목표
END_VAR
VAR_OUTPUT
	q_bNoCap	: BOOL;		// 용량·SOC 무효
END_VAR
VAR
	nMin		: UINT;
	fE			: REAL;		// kWh
END_VAR
M_AutoChg	:= 0.0;
q_bNoCap	:= i_stView.stGroup.fCapacity <= 0.0 OR NOT i_stView.stGroup.stSocAvg.bValid;
IF NOT q_bNoCap THEN
	nMin	:= F_MinutesTo(i_nNow := F_TimeHhmm(i_stTime := i_stView.stTime), i_nEnd := i_stWin.nEnd);
	fE		:= i_stView.stGroup.fCapacity * (i_stWin.fSoc - i_stView.stGroup.stSocAvg.fValue) / 100.0;
	IF nMin > 0 AND fE > 0.0 THEN
		M_AutoChg := MIN(MAX(fE * 60.0 / UINT_TO_REAL(nMin) + 1.0, 10.0), i_stView.stGroup.fPRatedAvail);
	END_IF
END_IF
END_METHOD

METHOD PROTECTED M_CheckTable : WSTRING(63)		// 시간표 칸 시각 점검 (시작 ≤ 끝, HHMM)
VAR_IN_OUT CONSTANT
	iq_stTable	: ST_CmScheduleSet;
END_VAR
VAR
	nS	: UINT;		// 계절
	nD	: UINT;		// 요일
	nK	: UINT;		// 칸
END_VAR
M_CheckTable := "";
FOR nS := 0 TO 2 DO
	FOR nD := 0 TO 6 DO
		FOR nK := 1 TO GVL_PARAM.SCHED_SLOT_COUNT DO
			IF NOT F_RealOk(iq_stTable.astSlot[nS, nD, nK].fP) THEN	// [결함 13 수정 2026-11-04: 칸 출력 kW가 숫자가 아님]
				M_CheckTable := WCONCAT(WCONCAT(WCONCAT(WCONCAT(WCONCAT("시간표 칸 출력 숫자 아님: 계절 ", TO_WSTRING(nS)), " 요일 "), TO_WSTRING(nD)), " 칸 "), TO_WSTRING(nK));
				RETURN;
			END_IF
			IF NOT F_HhmmOk(i_nHhmm := iq_stTable.astSlot[nS, nD, nK].nStart) OR NOT F_HhmmOk(i_nHhmm := iq_stTable.astSlot[nS, nD, nK].nEnd)
				OR iq_stTable.astSlot[nS, nD, nK].nStart > iq_stTable.astSlot[nS, nD, nK].nEnd THEN
				M_CheckTable := WCONCAT(WCONCAT(WCONCAT(WCONCAT(WCONCAT("시간표 칸 시각 잘못됨: 계절 ", TO_WSTRING(nS)), " 요일 "), TO_WSTRING(nD)), " 칸 "), TO_WSTRING(nK));
				RETURN;
			END_IF
		END_FOR
	END_FOR
END_FOR
END_METHOD

METHOD PROTECTED M_CheckWindow : BOOL		// 시간 구간 설정이 맞는가 (쓰지 않으면 TRUE)
VAR_INPUT
	i_stWin		: ST_CmWindowSet;
END_VAR
// [결함 13 수정 2026-11-04: SOC가 숫자가 아니면 (쓰지 않는 구간이어도) 틀림. 비교 전에 비트로. 원래 NOT i_stWin.bUse OR (… AND i_stWin.fSoc >= 0.0 AND i_stWin.fSoc <= 100.0)]
IF NOT F_RealOk(i_stWin.fSoc) THEN
	M_CheckWindow := FALSE;
	RETURN;
END_IF
M_CheckWindow := NOT i_stWin.bUse OR (F_HhmmOk(i_nHhmm := i_stWin.nStart) AND F_HhmmOk(i_nHhmm := i_stWin.nEnd)
	AND i_stWin.nStart <> i_stWin.nEnd AND i_stWin.fSoc >= 0.0 AND i_stWin.fSoc <= 100.0);
END_METHOD

METHOD M_ReasonText : WSTRING(63)
VAR_INPUT
	i_nReason	: UINT;
END_VAR
CASE i_nReason OF
	GVL_CM_RSN.NO_TIME:		M_ReasonText := "시각 무효";
	GVL_CM_RSN.NO_UNIT:		M_ReasonText := "가용 유닛 없음";
	GVL_CM_RSN.HOLIDAY:		M_ReasonText := "휴일";
	GVL_CM_RSN.NO_SLOT:		M_ReasonText := "맞는 시간표 칸 없음";
	GVL_CM_RSN.DIS_TIME:	M_ReasonText := "방전 허용 시간 아님";
	GVL_CM_RSN.REV_LIMIT:	M_ReasonText := "역송 방지로 방전 줄임";
	GVL_CM_RSN.NO_PCC:		M_ReasonText := "접속점 계측 무효 (방전 0)";
	GVL_CM_RSN.NO_CAP:		M_ReasonText := "배터리 용량·SOC 무효";
	GVL_CM_RSN.PEAK:		M_ReasonText := "피크 제어 방전";
	GVL_CM_RSN.BELOW_PEAK:	M_ReasonText := "피크 제어 필요 없음";
	GVL_CM_RSN.AUTO_CHG:	M_ReasonText := "자동 충전 시간";
	GVL_CM_RSN.REMAIN_DIS:	M_ReasonText := "잔량 방전 시간";
	GVL_CM_RSN.SCHED_PEAK:	M_ReasonText := "스케줄·피크 제어 중 큰 방전";
	GVL_CM_RSN.NEW_INTERVAL:	M_ReasonText := "새 15분 구간 시작";
ELSE
	M_ReasonText := WCONCAT("이유 ", TO_WSTRING(i_nReason));
END_CASE
END_METHOD

METHOD M_CheckSet : WSTRING(63)		// 공통 설정 점검. 파생 FB는 SUPER^.M_CheckSet() 뒤에 자기 설정을 점검
VAR
	k	: UINT;
END_VAR
M_CheckSet := "";
FOR k := 1 TO 12 DO
	IF i_stCommon.anSeasonOfMonth[k] > 2 THEN
		M_CheckSet := "제어 모드 공통: 월 → 계절 값은 0~2";
		RETURN;
	END_IF
END_FOR
IF NOT F_HhmmOk(i_nHhmm := i_stCommon.stDis.nStart) OR NOT F_HhmmOk(i_nHhmm := i_stCommon.stDis.nEnd) THEN
	M_CheckSet := "제어 모드 공통: 방전 허용 시간 HHMM";
ELSIF NOT (F_RealOk(i_stCommon.stNoRev.fMargin) AND F_RealOk(i_stCommon.stNoRev.fScale)) THEN	// [결함 13 수정 2026-11-04]
	M_CheckSet := "제어 모드 공통: 역송 방지 값 숫자 아님";
ELSIF i_stCommon.stNoRev.fMargin < 0.0 OR i_stCommon.stNoRev.fScale < 0.0 OR i_stCommon.stNoRev.fScale > 1.0 THEN
	M_CheckSet := "제어 모드 공통: 역송 방지 여유 0 이상, 비율 0~1";
END_IF
END_METHOD

END_FUNCTION_BLOCK

// ---- 10_Core/03_Base/FB_CtrlModeBase.TcPOU
FUNCTION_BLOCK ABSTRACT FB_CtrlModeBase EXTENDS FB_ModuleBase IMPLEMENTS I_ControlMode	// 제어 모드 공통 바탕. 파생 FB는 M_Calc만 쓰면 됨 (필요하면 M_CheckEnter·M_Enter·M_Exit·M_ReasonText·M_CheckSet을 바꿈)
// M_Enter·M_Exit를 바꾸면 SUPER^.M_Enter(i_stView := i_stView)·SUPER^.M_Exit()도 부름 (_bActive 유지)
VAR
	_bActive	: BOOL;		// 켜져 있음 (M_Enter ~ M_Exit). 진단용
END_VAR

METHOD M_CheckEnter : UINT		// 기본: 조건 없음
VAR_INPUT
	i_stView	: ST_CtrlModeView;	// 그룹 값(stGroup)·현지 시각(stTime). 관리자가 매 스캔 채움
END_VAR
M_CheckEnter := 0;
END_METHOD

METHOD M_Enter
VAR_INPUT
	i_stView	: ST_CtrlModeView;	// 그룹 값(stGroup)·현지 시각(stTime). 관리자가 매 스캔 채움
END_VAR
_bActive := TRUE;
END_METHOD

METHOD ABSTRACT M_Calc : ST_CtrlModeOut
VAR_INPUT
	i_stView	: ST_CtrlModeView;	// 그룹 값(stGroup)·현지 시각(stTime). 관리자가 매 스캔 채움
END_VAR
END_METHOD

METHOD M_Exit
_bActive := FALSE;
END_METHOD

END_FUNCTION_BLOCK

// ---- 10_Core/02_Util/F_InHhmmWindow.TcPOU
FUNCTION F_InHhmmWindow : BOOL		// 지금이 시간 구간 안인가: 시작 ≤ 지금 < 끝 (HHMM). 시작 > 끝이면 자정을 넘는 구간, 시작 = 끝이면 빈 구간
VAR_INPUT
	i_nNow		: UINT;		// HHMM
	i_nStart	: UINT;
	i_nEnd		: UINT;
END_VAR

IF i_nStart = i_nEnd THEN
	F_InHhmmWindow := FALSE;
ELSIF i_nStart < i_nEnd THEN
	F_InHhmmWindow := i_nNow >= i_nStart AND i_nNow < i_nEnd;
ELSE
	F_InHhmmWindow := i_nNow >= i_nStart OR i_nNow < i_nEnd;
END_IF

END_FUNCTION

// ---- 10_Core/02_Util/F_TimeHhmm.TcPOU
FUNCTION F_TimeHhmm : UINT		// 현지 시각 → HHMM (예: 13시 5분 = 1305)
VAR_INPUT
	i_stTime	: ST_LocalTime;
END_VAR

F_TimeHhmm := i_stTime.nHour * 100 + i_stTime.nMinute;

END_FUNCTION

// ---- 10_Core/02_Util/F_MinutesTo.TcPOU
FUNCTION F_MinutesTo : UINT		// 지금(HHMM)부터 끝(HHMM)까지 남은 분. 끝이 지났으면 다음 날 그 시각까지 (자정을 넘김). 같으면 0
VAR_INPUT
	i_nNow		: UINT;		// HHMM
	i_nEnd		: UINT;		// HHMM (2400 = 자정)
END_VAR
VAR
	nDiff		: DINT;
END_VAR

nDiff := (UINT_TO_DINT(i_nEnd / 100) * 60 + UINT_TO_DINT(i_nEnd MOD 100)) - (UINT_TO_DINT(i_nNow / 100) * 60 + UINT_TO_DINT(i_nNow MOD 100));
IF nDiff < 0 THEN
	nDiff := nDiff + 1440;
END_IF
F_MinutesTo := DINT_TO_UINT(nDiff);

END_FUNCTION

// ---- 10_Core/02_Util/F_HhmmOk.TcPOU
FUNCTION F_HhmmOk : BOOL		// HHMM 값이 맞는가: 0000~2359, 또는 2400 (하루 끝)
VAR_INPUT
	i_nHhmm		: UINT;
END_VAR

F_HhmmOk := ((i_nHhmm / 100) < 24 AND (i_nHhmm MOD 100) < 60) OR i_nHhmm = 2400;

END_FUNCTION

// ---- 20_Module/ControlMode/FB_CmConstPower.TcPOU
FUNCTION_BLOCK FB_CmConstPower EXTENDS FB_CtrlModeBase		// 제어 모드 예: 정출력. 설정한 P(·Q)를 접속점 기준으로 냄. tDuration이 지나면 스스로 끝냄
// 새 제어 모드의 본보기: FB_CtrlModeBase 상속 → M_Calc (+ 필요하면 M_CheckEnter·M_Enter·M_Exit·M_ReasonText·M_CheckSet)
VAR_INPUT
	i_stSet		: ST_CmConstPowerSet;	// 설정 (A_PassModuleSet이 GVL_PERSIST.g_stModuleSet 칸을 매 스캔 넘김)
END_VAR
VAR
	_tonRun		: TON;		// 운전 시간
END_VAR
VAR CONSTANT
	RSN_NO_UNIT	: UINT := 1;	// 진입 거부: 가용 유닛 없음
	RSN_TIME_UP	: UINT := 2;	// 끝: 운전 시간 끝
END_VAR

METHOD M_CheckEnter : UINT
VAR_INPUT
	i_stView	: ST_CtrlModeView;	// 그룹 값(stGroup)·현지 시각(stTime). 관리자가 매 스캔 채움
END_VAR
M_CheckEnter := 0;
IF i_stView.stGroup.nUnitAvail = 0 THEN
	M_CheckEnter := RSN_NO_UNIT;
END_IF
END_METHOD

METHOD M_Enter
VAR_INPUT
	i_stView	: ST_CtrlModeView;	// 그룹 값(stGroup)·현지 시각(stTime). 관리자가 매 스캔 채움
END_VAR
SUPER^.M_Enter(i_stView := i_stView);
_tonRun(IN := FALSE);		// 운전 시간을 처음부터 셈
END_METHOD

METHOD M_Calc : ST_CtrlModeOut
VAR_INPUT
	i_stView	: ST_CtrlModeView;	// 그룹 값(stGroup)·현지 시각(stTime). 관리자가 매 스캔 채움
END_VAR
_tonRun(IN := i_stSet.tDuration > T#0S, PT := i_stSet.tDuration);
M_Calc.bPSetActive	:= TRUE;
M_Calc.fPSet		:= i_stSet.fPSet;
M_Calc.bQSetActive	:= i_stSet.bQSet;
M_Calc.fQSet		:= i_stSet.fQSet;
M_Calc.bExitReq		:= FALSE;
M_Calc.nReason		:= 0;
IF _tonRun.Q THEN
	M_Calc.bExitReq	:= TRUE;
	M_Calc.nReason	:= RSN_TIME_UP;
END_IF
END_METHOD

METHOD M_CheckSet : WSTRING(63)		// 설정 점검: P·Q가 숫자인지 [결함 13 수정 2026-11-04: 추가. 원래 이 FB에는 점검 없음(바탕 FB 빈 문구)]
M_CheckSet := SUPER^.M_CheckSet();
IF M_CheckSet = "" AND NOT (F_RealOk(i_stSet.fPSet) AND F_RealOk(i_stSet.fQSet)) THEN
	M_CheckSet := "정출력: P·Q 값 숫자 아님";
END_IF
END_METHOD

METHOD M_ReasonText : WSTRING(63)
VAR_INPUT
	i_nReason	: UINT;
END_VAR
CASE i_nReason OF
	RSN_NO_UNIT:	M_ReasonText := "정출력: 가용 유닛 없음";
	RSN_TIME_UP:	M_ReasonText := "정출력: 운전 시간 끝";
ELSE
	M_ReasonText := WCONCAT("이유 ", TO_WSTRING(i_nReason));
END_CASE
END_METHOD

END_FUNCTION_BLOCK

// ---- 99_Test/PRG_TestSchedLive.TcPOU
PROGRAM PRG_TestSchedLive		// 스케줄 모드 실제 경로 시험 (시험 모드, MAIN이 부름): 지금 PLC 시각으로 시간표를 넣고 Auto → 배터리 투입 → Run → 스케줄 모드
// bStart := TRUE로 시작. 충전 칸 -200 kW (지금 분 ~ +2분) → 방전 칸 +100 kW (+2 ~ +4분) → 칸 없음 0 kW. 구간마다 5 s 안정 뒤 가상 PCS 실제 출력을 판정
// PCS1(유닛 1, 관리자 g_fbCtrlMode1)로 시험. 접속점은 실측 그대로(ePccShare := Actual)로 둠 (PCS2는 Manual 0)
// 시험 동안만: 방전 허용 시간 끔 (PLC 시계가 UTC), 가상신호로 수전 500 kW (가상 계측기는 부하가 없어 역송 방지에 걸림). 끝나면 설정·모드를 되돌리고 PCS 정지
VAR
	bStart		: BOOL;				// TRUE로 쓰면 시작 (시작하면 FALSE로 돌아감)
	bDone		: BOOL;				// 끝 (bPass로 결과)
	bPass		: BOOL;				// 세 구간 모두 맞음
	nStep		: UINT;
	wsStep		: WSTRING(80);		// 지금 단계
	wsFail		: WSTRING(80);		// 실패 이유
	(* 넣은 시간표 *)
	nSeason		: UINT;				// 0 여름, 1 봄·가을, 2 겨울
	nDow		: UINT;				// 0 = 일요일
	nChgStart	: UINT;				// HHMM, 충전 칸 시작
	nChgEnd		: UINT;				// HHMM, 충전 칸 끝 = 방전 칸 시작
	nDisEnd		: UINT;				// HHMM, 방전 칸 끝
	(* 지금 값 *)
	stNow		: ST_LocalTime;		// PLC 시각 (MAIN.fbClock)
	nActiveMode	: UINT;				// 관리자 켜진 모드 (2 = 스케줄)
	nSlot		: UINT;				// 스케줄 모드가 맞춘 칸
	nSchedState	: UINT;				// 스케줄 모드 상태 (GVL_CM_RSN)
	fSchedP		: REAL;				// 스케줄 모드가 낸 값 (kW, 방전 +)
	fMgrP		: REAL;				// 관리자 지령 (지령원 출력, kW)
	fUnitP		: REAL;				// 가상 PCS 실제 출력 (kW, 방전 +)
	eRun		: E_RunState;		// 가상 PCS 운전 상태
	(* 판정: 구간마다 안정 뒤 값 *)
	fChgP		: REAL;
	fDisP		: REAL;
	fZeroP		: REAL;
	bChgOk		: BOOL;
	bDisOk		: BOOL;
	bZeroOk		: BOOL;
	(* 내부 *)
	nLastStep	: UINT;
	tonStep		: TON;				// 단계 시간 초과
	tonSettle	: TON;				// 구간 진입 뒤 안정
	bBackedUp	: BOOL;
	stSchedBak	: ST_CmScheduleSet;
	stCommonBak	: ST_CmCommonSet;
	stCmBak		: ST_CtrlModeSet;
	stVirtBak	: ST_VirtualSet;
	stMgrOut	: ST_SourceOutput;
	nMin		: UINT;
	k			: UINT;
END_VAR

// 지금 값 (화면용)
stNow		:= MAIN.fbClock.q_stTime;
nActiveMode	:= GVL_SITE.g_fbCtrlMode1.q_nActive;
nSlot		:= GVL_SITE.g_fbCmSchedule1.q_nSlot;
nSchedState	:= GVL_SITE.g_fbCmSchedule1.q_nState;
fSchedP		:= GVL_SITE.g_fbCmSchedule1.q_fOutP;
stMgrOut	:= GVL_SITE.g_fbCtrlMode1.Output;
fMgrP		:= stMgrOut.fPSet;	// [16번 수정 2026-11-09: 관리자가 접속점 그룹 단위 → 접속점 그룹 지령 칸. 원래 stMgrOut.astUnit[1].fPSet (PCS2는 Manual이라 접속점 그룹 지령이 유닛 1로 감)]
fUnitP		:= MAIN.fbSnapshot.q_astUnit[1].stP.fValue;
eRun		:= MAIN.fbSnapshot.q_astUnit[1].eRunState;

tonStep(IN := nStep >= 20 AND nStep < 90, PT := T#200S);

CASE nStep OF
	0:
		IF bStart THEN
			bStart		:= FALSE;
			bDone		:= FALSE;
			bPass		:= FALSE;
			bChgOk		:= FALSE;
			bDisOk		:= FALSE;
			bZeroOk		:= FALSE;
			fChgP		:= 0.0;
			fDisP		:= 0.0;
			fZeroP		:= 0.0;
			wsFail		:= "";
			nStep		:= 10;
		ELSIF NOT bDone THEN
			wsStep := "대기: bStart := TRUE로 시작";
		END_IF

	10:	// 지금 시각으로 시간표 넣기
		wsStep := "시간표 넣는 중";
		IF NOT stNow.bValid OR stNow.nMonth < 1 OR stNow.nMonth > 12 OR stNow.nDay < 1 OR stNow.nDay > 31 OR stNow.nDayOfWeek > 6 THEN
			wsFail	:= "PLC 시각 무효";
			nStep	:= 90;
		ELSE
			nMin := stNow.nHour * 60 + stNow.nMinute;
			IF nMin + 4 >= 1440 THEN
				wsFail	:= "자정 직전이라 시험 안 함 (몇 분 뒤 다시)";
				nStep	:= 90;
			ELSE
				stSchedBak	:= GVL_PERSIST.g_stModuleSet.stCmSchedule1;
				stCommonBak	:= GVL_PERSIST.g_stModuleSet.stCmCommon;
				stVirtBak	:= GVL_TEST.g_astVirtual[1];
				stCmBak		:= GVL_PERSIST.g_stModuleSet.stCtrlMode1;
				GVL_PERSIST.g_stModuleSet.stCtrlMode1.ePccShare := E_PccShare.Actual;
				bBackedUp	:= TRUE;
				nSeason := GVL_PERSIST.g_stModuleSet.stCmCommon.anSeasonOfMonth[stNow.nMonth];
				IF nSeason > 2 THEN
					nSeason := 0;
				END_IF
				nDow		:= stNow.nDayOfWeek;
				nChgStart	:= (nMin / 60) * 100 + nMin MOD 60;
				nChgEnd		:= ((nMin + 2) / 60) * 100 + (nMin + 2) MOD 60;
				nDisEnd		:= ((nMin + 4) / 60) * 100 + (nMin + 4) MOD 60;
				FOR k := 1 TO GVL_PARAM.SCHED_SLOT_COUNT DO
					GVL_PERSIST.g_stModuleSet.stCmSchedule1.astSlot[nSeason, nDow, k].nStart	:= 0;
					GVL_PERSIST.g_stModuleSet.stCmSchedule1.astSlot[nSeason, nDow, k].nEnd	:= 0;
					GVL_PERSIST.g_stModuleSet.stCmSchedule1.astSlot[nSeason, nDow, k].fP		:= 0.0;
				END_FOR
				GVL_PERSIST.g_stModuleSet.stCmSchedule1.astSlot[nSeason, nDow, 1].nStart	:= nChgStart;
				GVL_PERSIST.g_stModuleSet.stCmSchedule1.astSlot[nSeason, nDow, 1].nEnd	:= nChgEnd;
				GVL_PERSIST.g_stModuleSet.stCmSchedule1.astSlot[nSeason, nDow, 1].fP		:= -200.0;
				GVL_PERSIST.g_stModuleSet.stCmSchedule1.astSlot[nSeason, nDow, 2].nStart	:= nChgEnd;
				GVL_PERSIST.g_stModuleSet.stCmSchedule1.astSlot[nSeason, nDow, 2].nEnd	:= nDisEnd;
				GVL_PERSIST.g_stModuleSet.stCmSchedule1.astSlot[nSeason, nDow, 2].fP		:= 100.0;
				GVL_PERSIST.g_stModuleSet.stCmCommon.abHoliday[stNow.nMonth, stNow.nDay]	:= FALSE;
				GVL_PERSIST.g_stModuleSet.stCmCommon.stDis.bUse	:= FALSE;
				GVL_TEST.g_astVirtual[1].bPEna	:= TRUE;
				GVL_TEST.g_astVirtual[1].fP		:= -500.0;		// 수전 500 kW
				GVL_PERSIST.g_aeOpMode[1]		:= E_OpMode.Auto;
				nStep := 20;
			END_IF
		END_IF

	20:	// Auto 전환 → 배터리 투입 요청
		wsStep := "Auto 전환 대기";
		IF MAIN.fbModeSwitch.q_aeOpMode[1] = E_OpMode.Auto THEN
			GVL_SITE.g_fbSrcTest.i_nBatGroup	:= 0;
			GVL_SITE.g_fbSrcTest.i_eBatReq		:= E_BatCmd.Close;
			nStep := 30;
		END_IF

	30:	// 배터리 투입 → Run 요청
		wsStep := "배터리 투입 대기";
		IF MAIN.fbBatGroup.q_astBatGroup[1].bReady THEN
			GVL_SITE.g_fbSrcTest.i_nPcsUnit	:= 0;
			GVL_SITE.g_fbSrcTest.i_ePcsReq	:= E_PcsCmd.Run;
			nStep := 40;
		END_IF

	40:	// Run → 스케줄 모드(2) 요청
		wsStep := "PCS Run 대기";
		IF eRun = E_RunState.Run THEN
			GVL_SITE.g_fbCtrlMode1.i_nModeReq := 2;
			nStep := 50;
		END_IF

	50:
		wsStep := "스케줄 모드 켜는 중";
		IF nActiveMode = 2 THEN
			nStep := 60;
		END_IF

	60:	// 충전 칸
		wsStep := "충전 칸: -200 kW";
		tonSettle(IN := nSlot = 1, PT := T#5S);
		IF tonSettle.Q THEN
			fChgP	:= fUnitP;
			bChgOk	:= ABS(fUnitP + 200.0) < 5.0 AND ABS(fSchedP + 200.0) < 0.1 AND ABS(fMgrP + 200.0) < 0.1;
		END_IF
		IF nSlot = 2 THEN
			tonSettle(IN := FALSE);
			nStep := 70;
		END_IF

	70:	// 방전 칸
		wsStep := "방전 칸: +100 kW";
		tonSettle(IN := nSlot = 2, PT := T#5S);
		IF tonSettle.Q THEN
			fDisP	:= fUnitP;
			bDisOk	:= ABS(fUnitP - 100.0) < 5.0 AND ABS(fSchedP - 100.0) < 0.1 AND ABS(fMgrP - 100.0) < 0.1;
		END_IF
		IF nSlot = 0 THEN
			tonSettle(IN := FALSE);
			nStep := 80;
		END_IF

	80:	// 칸 없음 → 0
		wsStep := "칸 없음: 0 kW";
		tonSettle(IN := nSlot = 0, PT := T#5S);
		IF tonSettle.Q THEN
			fZeroP	:= fUnitP;
			bZeroOk	:= ABS(fUnitP) < 5.0 AND nSchedState = GVL_CM_RSN.NO_SLOT AND stMgrOut.bPSetActive;	// [16번 수정 2026-11-09: 원래 stMgrOut.astUnit[1].bPSetActive]
			tonSettle(IN := FALSE);
			nStep := 90;
		END_IF

	90:	// 정리: 모드 끔, PCS 정지, 설정·가상신호·운전 모드 되돌림
		GVL_SITE.g_fbCtrlMode1.i_nModeReq	:= 0;
		GVL_SITE.g_fbSrcTest.i_nPcsUnit		:= 0;
		GVL_SITE.g_fbSrcTest.i_ePcsReq		:= E_PcsCmd.Stop;
		IF bBackedUp THEN
			GVL_PERSIST.g_stModuleSet.stCmSchedule1	:= stSchedBak;
			GVL_PERSIST.g_stModuleSet.stCmCommon	:= stCommonBak;
			GVL_TEST.g_astVirtual[1]				:= stVirtBak;
			GVL_PERSIST.g_stModuleSet.stCtrlMode1	:= stCmBak;
			bBackedUp := FALSE;
		END_IF
		GVL_PERSIST.g_aeOpMode[1] := E_OpMode.Manual;
		bPass	:= bChgOk AND bDisOk AND bZeroOk AND wsFail = "";
		bDone	:= TRUE;
		IF bPass THEN
			wsStep := "끝: 통과";
		ELSE
			wsStep := "끝: 실패 (wsFail·구간 값 확인)";
		END_IF
		nStep := 0;
END_CASE

// 단계 시간 초과
IF tonStep.Q AND nStep >= 20 AND nStep < 90 THEN
	wsFail	:= WCONCAT("시간 초과: ", wsStep);
	nStep	:= 90;
END_IF
IF nStep <> nLastStep THEN
	tonStep(IN := FALSE);
	nLastStep := nStep;
END_IF

END_PROGRAM

